(* IEC 61131-3 sources: JingjiangMoonbox/Application/Application/数据类型/系统参数/保持参数, 3 files *)

(* ---- StGrpParam_Save.st ---- *)
(*@CES
Name=StGrpParam_Save
Type=Gvl
TypeGuid=2db5746d-d284-4425-9f7f-2663a34b0ebc
Guid=f58940ec-a17f-4bea-a7e2-f076956df0df
HasDeclaration=True
HasImplementation=False
*)
{DECLARATION}
{attribute 'pack_mode' := '1'}
TYPE StGrpParam_Save :
STRUCT
	rGirth_BottomRoller							: REAL;(* 底辊周长/整机设置状态 *)
	uiNum_BottomRoller							: UINT;(* 底辊减速比分子/整机设置状态 *)
	uiDen_BottomRoller							: UINT;(* 底辊减速比分母/整机设置状态 *)

	rGirth_PrnRoller							: REAL;(* 印版周长/整机设置状态 *)
	uiNum_PrnRoller								: UINT;(* 版辊减速比分子/整机设置状态 *)
	uiDen_PrnRoller								: UINT;(* 版辊减速比分母/整机设置状态 *)

	rGirth_NetRoller							: REAL;(* 网辊周长/整机设置状态 *)
	uiNum_NetRoller								: UINT;(* 网辊减速比分子/整机设置状态 *)
	uiDen_NetRoller								: UINT;(* 网辊减速比分母/整机设置状态 *)

	rGirth_StrRoller							: REAL;(* 张带辊周长 *)
	uiNum_StrRoller								: UINT;(* 张带辊减速比分子/整机设置状态 *)
	uiDen_StrRoller								: UINT;(* 张带辊减速比分母/整机设置状态 *)

	rScrewPitch_PrnRoller_Pressure				: REAL;(* 版辊压力架丝杆节距/整机设置状态/单位mm *)
	uiNum_PrnRoller_Pressure					: UINT;(* 版辊压力电机减速比分子/整机设置状态 *)
	uiDen_PrnRoller_Pressure					: UINT;(* 版辊压力电机减速比分母/整机设置状态 *)

	rScrewPitch_NetRoller_Pressure				: REAL;(* 网辊压力架丝杆节距/整机设置状态/单位mm *)
	uiNum_NetRoller_Pressure					: UINT;(* 网辊压力电机减速比分子/整机设置状态 *)
	uiDen_NetRoller_Pressure					: UINT;(* 网辊压力电机减速比分母/整机设置状态 *)

	rScrewPitch_StrRoller_Pressure				: REAL;(* 张带辊压力架丝杆节距/整机设置状态/单位mm *)
	uiNum_StrRoller_Pressure					: UINT;(* 张带辊压力电机减速比分子/整机设置状态 *)
	uiDen_StrRoller_Pressure					: UINT;(* 张带辊压力电机减速比分母/整机设置状态 *)

	rGirth_CenterRoller							: REAL;(* 中心辊周长/整机设置状态 *)
	uiNum_CenterRoller							: UINT;(* 中心辊减速比分子/整机设置状态 *)
	uiDen_CenterRoller							: UINT;(* 中心辊减速比分母/整机设置状态 *)

	rScrewPitch_Horz							: REAL;(* 横向架丝杆节距/整机设置状态/单位mm *)
	uiNum_Horz									: UINT;(* 横向电机减速比分子/整机设置状态 *)
	uiDen_Horz									: UINT;(* 横向电机减速比分母/整机设置状态 *)

	rScrewPitch_PhotoCell						: REAL;(* 光电眼架丝杆节距/整机设置状态/单位mm *)
	uiNum_PhotoCell								: UINT;(* 光电眼电机减速比分子/整机设置状态 *)
	uiDen_PhotoCell								: UINT;(* 光电眼电机减速比分母/整机设置状态 *)

	wAI_polarity								: WORD;(* 模拟量输入极性配置 *)
		(*
		/bit0=1放料模拟量输入反向
		/bit1=1收料模拟量输入反向
		/bit2=1放牵模拟量输入反向
		/bit3=1收牵模拟量输入反向
		/bit4~bit15(保留)
		/ *)
	lrPrnLen_AmountTo							: LREAL;(* 总计印刷长度/单位:m *)
	rPrintLengthCoef							: REAL;(*印刷计长系数|*)
	alrPrnLen									: ARRAY [1..3] OF LREAL;(* A轴印长/B轴印长/总印长 *)
	alrPrnLen_Alr								: ARRAY [1..3] OF LREAL;(* 印长报警值/相对应于alrPrnLen *)
	iDelayMsec_RollerPress						: INT;(* 压辊延时/单位:ms *)

	wUwRwAxisProf								: WORD;
(*												/放料&收料轴描述 *)
(*												/bit0=TRUE,放料当前轴A轴 *)
(*												/bit1=TRUE,收料当前轴A轴 *)

	iMarkTypeId									: INT;(* 色标形式 *)
	iMarkArrangeMode							: INT;(* 标记排列形式 *)
	byTriMark_SideC								: BYTE;(* 梯形色标直边(c边) *)
	byTriMark_SideB								: BYTE;(* 梯形色标底边(b边) *)
	bySysSamplePrecision						: BYTE;(*系统采样精度			*)
	byArcFineSampleType							: BYTE;(*系统采样方式*)

	(* 时间设定 *)
	iTime_Stop									: INT;(* 停机时间/单位:s *)
	iTime_Estop									: INT;(* 急停时间/单位:s *)
	iTime_AutoAcc							: INT;(* 自动加减速时间/单位:s *)
	iTime_ManuAcc							: INT;(* 手动加减速时间/单位:s *)
	iTime_S										: INT;(* S加减速时间/单位:s *)
	iTime_PreDrvAcc_Uw								: INT;(* 预驱加速时间/10s *)
	iTime_PreDrvDec_Uw							: INT;(* 预驱减速时间/2s *)
	iTime_PreDrvAcc_Rw								: INT;(* 预驱加速时间/10s *)
	iTime_PreDrvDec_Rw							: INT;(* 预驱减速时间/2s *)
	iTime_FilmAcc								: INT;(* 料膜加速时间/8S *)
	iTime_FilmDec								: INT;(* 料膜减速时间/2S *)
	iTime_AutoDec							: INT;(*自动加减速时间|单位:s|*)
	iTime_ManuDec							: INT;(*手动加减速时间|单位:s|*)
	iTime_FastStop							: INT;(*快停时间*)
	iTime_S_End								: INT;(*S减加速时间*)
	byAutoAccDecCurve					: BYTE;(*自动加减速曲线选择|默认 按照最大直线加速度进行s处理-
																		 1：按照直线加速时间进行s处理
																		 2：按照直线加速时间全程s处理-*)

	rVel_Max									: REAL;(* 设备最大速度/单位:m/min *)
	rVel_Tar									: REAL;(* 目标速度/单位:m/min *)
	arVel_Usr									: ARRAY [1..3] OF REAL;(* 用户速度1,2,3/单位:m/min *)
	rVel_Ink									: REAL;(* 匀墨速度/单位:m/min *)
	rVel_Inch									: REAL;(* 单运行速度/单位:m/min *)
	rVel_AutoAdj								: REAL;(* 自动修正速度/单位:m/min *)
	rVel_ManuAdj_Corse							: REAL;(* 手动粗调速度/单位:m/min *)
	rVel_ManuAdj_Fine							: REAL;(* 手动细调速度/单位:m/min *)
	rVel_RapidAdj								: REAL;(* 快速调版速度/单位:m/min *)
	rVel_HorzdAdj								: REAL;(* 横向调版速度/单位:mm/s *)

	rDiamAlarm_Uw								: REAL;(* 放料报警卷径 *)
	rGirth_AxiaA_Uw								: REAL;(* 放料A轴周长 *)
	rGirth_AxiaB_Uw								: REAL;(* 放料B轴周长 *)
	arKpid_Uw									: ARRAY [1..3] OF REAL;(* 放料pid比例 *)
	rGirth_Uw									: REAL;(* 放料周长 *)
	uiNum_Uw									: UINT;(* 放料减速比-电机转数 *)
	uiDen_Uw									: UINT;(* 放料减速比-负载转数 *)
	rTaper_Uw									: REAL;(* 放料锥度 *)
	rAI_med_Uw									: REAL;(* 放料摆臂模拟量中位 *)
	byDiamMeasureTypeId_Uw						: BYTE;(* 放料卷径测量类型 *)
	byAIType_Uw									: BYTE;(* 放料摆臂类型/初始值0 *)
	byCoef_stiffen_Uw							: BYTE;(* 放料拉料系数|10 *)

	adwEnc_AxisALocation_Uw						: ARRAY [0..1] OF DWORD;(* 放料A轴定位位置/索引通过BOOL_TO_INT(xCutterOnTop_#w)来访问 *)
	adwEnc_AxisALocation_MinDiam_Uw				: ARRAY [0..1] OF DWORD;(* 放料A轴最小径位置/索引通过BOOL_TO_INT(xCutterOnTop_#w)来访问 *)
	adwEnc_AxisBLocation_Uw						: ARRAY [0..1] OF DWORD;(* 放料B轴定位位置/索引通过BOOL_TO_INT(xCutterOnTop_#w)来访问 *)
	adwEnc_AxisBLocation_MinDiam_Uw				: ARRAY [0..1] OF DWORD;(* 放料B轴最小径位置/索引通过BOOL_TO_INT(xCutterOnTop_#w)来访问 *)
	iRatedRpm_Uw								: INT;(* 放料电机额定转速/1500r/min *)
	iRatedFreq_Uw								: INT;(* 放料电机额定频率/50HZ *)
	iUpperFreq_Uw								: INT;(* 放料电机上限频率/100HZ *)
	xDiamMeasureAutomatic_Uw					: BOOL;(* 放料卷径自动测量标志/FALSE *)
	xCutUseReflectionSensor_Uw					: BOOL;(* 放料采用弧面检测方式标志,TRUE标识有效/FALSE *)
	xMultAxisParaEn_Uw							: BOOL;(* 放料AB轴单独参数-卷径测量/FALSE *)
	xFlag_CCW_AfterCutted_Uw					: BOOL;(* 裁切后放料轴反转/TRUE *)
	iPreRevLenth_MM_Cutted_Uw					: INT;(* 放料轴裁切反转距离/初始值1000 *)
	iPreRevVel_RPM_Cutted_Uw					: INT;(* 放料轴裁切反转转速/初始值80 *)
	xPreCutOneBtn_Uw							: BOOL;(* 放料接料准备使用单输入标志/FALSE *)
	rCoefCut_FilmVolPerimeter_Uw				: REAL;(* 放料裁切系数/1.5 *)
	xDiaEstEn_Uw								: BOOL;(* 放料卷径估计使能/FALSE *)
	rEstiDia_Uw									: REAL;(* 预估卷径值/300mm *)
	rEstiThickness_Uw							: REAL;(* 预估料膜厚度值/0.02mm *)
	byDelayTime_DiaCompensateWhenCutDne_Uw		: BYTE;(* 裁切后卷径补偿介入时间/10s *)
	uiPiDelay_Uw								: UINT;(* 裁切后放料PI延迟时间/1000ms *)

	xUseRadCompensate_Uw						: BOOL;(* 放料翻转架补偿使能标志/FALSE *)
	xConfirmRad0_Uw								: BOOL;(* 放料确认弧度0标志/FALSE *)
	dwAxisAabsPos_0Rad_Uw						: DWORD;(* 放料A轴翻转架0度的绝对位置/翻转架中心作为坐标系0点/0 *)
	dwAxisBabsPos_0Rad_Uw						: DWORD;(* 放料B轴翻转架0度的绝对位置/翻转架中心作为坐标系0点/0 *)
	(*											/ALTMA的放料架结构 *)
	rDiam_Tower_Uw								: REAL;(* 放料翻转架的直径/1000mm *)
	rDiam_NextRoller_Uw							: REAL;(* 放料翻转架下个辊的直径/100mm *)
	rXPos_NextRoller_Uw							: REAL;(* 放料翻转架下个辊的X位置/232.5mm/翻转架中心作为坐标系0点 *)
	rYPos_NextRoller_Uw							: REAL;(* 放料翻转架下个辊的Y位置/1052mm/翻转架中心作为坐标系0点 *)
	xTowerDir_Uw								: BOOL;(* 翻转架和绝对位置方向控制/FALSE *)
	(*2022.5.17.121911 放料翻转架补偿算法优化后增加的变量|13bytes|2023.8.17.161013*)
	rDiam_DeflectorRollPos_Uw				: REAL;(*翻料架的导向辊圆心运动直径|距离翻转架圆心=该值/2|mm*)
	rDiam_DeflectorRoller_Uw				: REAL;(*翻料架上导向辊的直径|mm*)
	xMultAxisPosEn_Uw							: BOOL;(* 放料定位位置单独参数-绝对值编码器/FALSE *)
	byInitialSpd_Stiffen_Uw						: BYTE;(* 放料拉料初始速度/10r/min *)
	(*											/ 2021.11.5.174244 *)
	rFilmLen_UnwindToPU1						: REAL;(*放料裁切点到1U的料膜距离|单位:mm|*)
	rFilmLen_NotAdjFront						: REAL;(*裁切点前不调整的料长|单位:mm|*)
	rFilmLen_NotAdjBack							: REAL;(*裁切点后不调整的料长|单位:mm|*)
	rFilmLen_BetweenImpressPoints				: REAL;(*两个压印点之间的料长|单位:mm|*)

	rDiamAlarm_Rw								: REAL;(* 收料报警卷径 *)
	rGirth_AxiaA_Rw								: REAL;(* 收料A轴周长 *)
	rGirth_AxiaB_Rw								: REAL;(* 收料B轴周长 *)
	arKpid_Rw									: ARRAY [1..3] OF REAL;(* 放料pid比例 *)
	rGirth_Rw									: REAL;(* 收料周长 *)
	uiNum_Rw									: UINT;(* 收料减速比-电机转数 *)
	uiDen_Rw									: UINT;(* 收料减速比-负载转数 *)
	rAI_med_Rw									: REAL;(* 收料摆臂模拟量中位 *)
	byAIType_Rw									: BYTE;(* 收料摆臂类型/初始值0 *)
	byCoef_stiffen_Rw							: BYTE;(* 收料拉料系数|10 *)
	xRsv										: BOOL;
	adwEnc_AxisALocation_Rw						: ARRAY [0..1,0..1] OF DWORD;(* 收料A轴定位位置/一维索引通过BOOL_TO_INT(xCutterOnTop_Rw)/二维索引[0]表示3吋纸芯,[1]表示6吋纸芯 *)
	adwEnc_AxisBLocation_Rw						: ARRAY [0..1,0..1] OF DWORD;(* 收料B轴定位位置/一维索引通过BOOL_TO_INT(xCutterOnTop_Rw)/二维索引[0]表示3吋纸芯,[1]表示6吋纸芯 *)
	rTaper_begin_Rw								: REAL;(* 锥度起始值-收料 *)
	rTaper_end_Rw								: REAL;(* 锥度结束值-收料 *)
	rDiam_taper_begin_Rw						: REAL;(* 锥度起始直径-收料 *)
	rDiam_taper_end_Rw							: REAL;(* 锥度结束直径-收料 *)
	iRatedRpm_Rw								: INT;(* 收料电机额定转速/默认1500 *)
	iRatedFreq_Rw								: INT;(* 收料电机额定频率/默认50 *)
	iUpperFreq_Rw								: INT;(* 收料电机上限频率/默认100 *)
	rGirth_3inch_Rw								: REAL;(* 收料3寸周长/默认300 *)
	rGirth_6inch_Rw								: REAL;(* 收料6寸周长/默认600 *)
	xPreCutOneBtn_Rw							: BOOL;(* 收料接料准备使用单输入标志/默认FALSE *)
	rCoefCut_FilmVolPerimeter_Rw				: REAL;(* 收料裁切系数/0.5 *)
	xDiaEstEn_Rw								: BOOL;(* 收料卷径估计使能/默认FALSE *)
	rEstiDia_Rw									: REAL;(* 预估卷径值/默认300mm *)
	rEstiThickness_Rw							: REAL;(* 预估料膜厚度值/默认0.02mm *)
	byDelayTime_DiaCompensateWhenCutDne_Rw		: BYTE;(* 裁切后卷径补偿介入时间/默认10s *)
	xUseAbsEncEn_Rw								: BOOL;(* 收料使用绝对值编码器标志/默认FALSE *)
	xMultAxisPosEn_Rw							: BOOL;(* 收料定位位置单独参数-绝对值编码器/默认FALSE *)
	byInitialSpd_Stiffen_Rw						: BYTE;(* 收料拉料初始速度/10r/min *)

	rDiamCurAxis_Uw								: REAL;(* 放料当前卷径 *)
	rDiamCurAxis_Rw								: REAL;(* 收料当前卷径 *)

	rGirth_If									: REAL;(* 放牵周长 *)
	uiNum_If									: UINT;(* 放牵减速比-电机转数 *)
	uiDen_If									: UINT;(* 放牵减速比-负载转数 *)
	rTaper_If									: REAL;(* 放牵锥度 *)
	byAIType_If									: BYTE;(* 放牵摆臂类型/初始值0 *)
	rAI_med_If									: REAL;(* 放牵摆臂模拟量中位 *)
	arKpid_If									: ARRAY [1..3] OF REAL;(* 放牵pid/2021.11.18.201839 *)
	iRatedRpm_If								: INT;(* 放牵电机额定转速/1500rpm *)
	iRatedFreq_If								: INT;(* 放牵电机额定频率/50HZ *)
	iUpperFreq_If								: INT;(* 放牵电机上限频率/100HZ *)
	xInchNegative_If							: BOOL;(* 放牵单运行反向/FALSE *)
	iInchVel_If									: INT;(* 放牵单运行速度/10m/min *)

	rGirth_Of									: REAL;(* 收牵周长 *)
	uiNum_Of									: UINT;(* 收牵减速比-电机转数 *)
	uiDen_Of									: UINT;(* 收牵减速比-负载转数 *)
	rTaper_Of									: REAL;(* 收牵锥度 *)
	byAIType_Of									: BYTE;(* 收牵摆臂类型/初始值0 *)
	rAI_med_Of									: REAL;(* 收牵摆臂模拟量中位 *)
	arKpid_Of									: ARRAY [1..3] OF REAL;(* 收牵pid/2021.11.18.202112 *)
	iRatedRpm_Of								: INT;(* 收牵电机额定转速/1500rpm *)
	iRatedFreq_Of								: INT;(* 收牵电机额定频率/50HZ *)
	iUpperFreq_Of								: INT;(* 收牵电机上限频率/100HZ *)
	xInchNegative_Of							: BOOL;(* 收牵单运行反向/FALSE *)
	iInchVel_Of									: INT;(* 收牵单运行速度/10m/min *)

(*2025.8.4.144213|原dwExtBitCtlFlag变量-改为BIT型--*)
	xSwitch_Change_CutterOnTop_HMI_Uw			: BIT;(*放料上下裁切换-界面按钮bit2*)
	xSwitch_Change_CutterOnTop_HMI_Rw			: BIT;(*收料上下裁切换-界面按钮bit3*)
	xCancelTenEn								: BIT;(*取消张力规划使能开bit10*)
	xEn_DualParam_AbsEncLocation_Uw				: BIT;(*bit11: 放料编码器方式下定位使用多轴使能|2021.5.7.111434|Liu.yt*)
	xEn_DualParam_AbsEncLocation_Rw				: BIT;(*bit12: 收料编码器方式下定位使用多轴使能|2021.5.7.111434|Liu.yt*)
	xFlag_AxisABParaFroDiaMea_Uw				: BIT;(*放料自动卷径分轴标志*)
	xSwitchTension_If							: BIT;(*bit6 放牵张力算法切换/FALSE *)
	xSwitchTension_Of							: BIT;(*bit7 收牵张力算法切换/FALSE *)
	xEnFeedLimitWarnFlag						: BIT;(*bit5 牵引速度限制提示使能位*)
	xSwitch_AxisLocaltion_DualParam_Uw			: BIT;(*放料绝对值编码器定位双轴参数开关|原bit11*)
	xSwitch_AxisLocaltion_DualParam_Rw			: BIT;(*收料绝对值编码器定位双轴参数开关|原bit12*)
	dwExtBitCtlFlag								: DWORD;(*扩展位控制标志|2019.1.25.143212|
													*.bit0: 放料自动卷径是否分轴来作?|FALSE默认一起|TRUE表示ab轴分开||
													*.bit1: 一键开机使能标志||
													*.bit2: 放料上下裁控制开关(区分于xCutterOnTop_Uw|)|2019.3.28.092931|补充遗漏||
													*.bit3: 收料上下裁控制开关(区分于xCutterOnTop_Rw|)|2019.3.28.092931|补充遗漏||
													Deprecated@2019.8.13.115259|*.bit4: 超声波检测使能|2019.3.23.154021||2019.3.28.092949|纠正错误||
													*.bit5: 牵引速度限制提示使能位|2019.4.18.135612|xie.gc||
													*.bit6: 放牵算法切换开关|@2019.8.1.091703|
													*.bit7: 收牵算法切换开关|@2019.8.1.091703|
													*.bit8: 放料前馈使能位|@2019.8.8.162527|xie.gc|
													*.bit9: 收料前馈使能位|@2019.8.8.162527|xie.gc|
													*.bit10: 取消张力规划使能开|2019.10.14.152513|niu.j|
													*.bit11: 放料编码器方式下定位使用多轴使能|2021.5.7.111434|Liu.yt|
													*.bit12: 收料编码器方式下定位使用多轴使能|2021.6.1.093832|Liu.yt|
													ALTMA增加了上下裁刀是否配置标志
													*.bit13: |2021.7.17.142536 放料上裁刀开启|Liu.yt|
													*.bit14: |2021.7.17.142536 放料下裁刀开启|Liu.yt|
													*.bit15: |2021.7.17.142536 收料上裁刀开启|Liu.yt|
													*.bit16: |2021.7.17.142536 收料下裁刀开启|Liu.yt|
													*.bit17: 2022.4.6.130956\翻料架打开控制位|
													|*)

	byTaperCtlMode_Uw							: BYTE;(*锥度调整方式*)
	byTaperCtlMode_Rw							: BYTE;(*锥度调整方式*)
	(*2022.4.14.094534 收放料自动接料|21BYTES*)
	xAutomaticCutEn_Uw							: BOOL;(*放料自动裁切使能|*)
	byAutoMaticCutMode_Uw						: BYTE;(*放料自动裁切模式|0 按照剩余米数
																	 |1 按照剩余卷径*)
	uiAutoMaticCutMeters_Uw						: UINT;(*自动裁切米数|m*)
	uiAutoMaticCutDia_Uw						: UINT;(*自动裁切卷径|*)

	xAutomaticCutEn_Rw							: BOOL;(*收料自动裁切使能|*)
	byAutoMaticCutMode_Rw						: BYTE;(*收料自动裁切模式|0 按照计米长度-在上次接料完成后启动
															         |1 按照放料裁切后整机长度-在放料接料完成后启动
																     |2 按照当前卷径-在上次接料完成后启动*)
	uiAutoMaticCutMeters_Rw						: UINT;(*自动裁切米数|m*)
	uiAutoMaticCutDia_Rw						: UINT;(*自动裁切卷径|*)
	byLenth_Machine								: BYTE;(*整机长度|m*)
	rDia_PaperRoller_Uw							: REAL;(*纸筒直径|mm*)
	rFilmThickNess								: REAL;(*料膜厚度|mm*)
	(*放料|*)
	rDiamTaper_Begin_Uw							: REAL;(*放料起始锥度对应卷径|*)
	rDiamTaper_End_Uw							: REAL;(*放料结束锥度对应卷径|*)
	rTaper_Begin_Uw								: REAL;(*锥度起始|放料|*)
	rTaper_End_Uw								: REAL;(*锥度结束|放料|*)

	(*放牵|*)
	rTaper_Begin_If								: REAL;(*锥度起始|放牵|*)
	rTaper_End_If								: REAL;(*锥度结束|放牵|*)
	(*收牵|*)
	rTaper_Begin_Of								: REAL;(*锥度起始|收牵|*)
	rTaper_End_Of								: REAL;(*锥度结束|收牵|*)

	xStep_Fast:BOOL;
	rStep_Fast:REAL;
	rStep_Little:REAL;
(*增加收放料收放牵锥度单位切换|支持%、N、mpa|104bytes*)
	byTaperUnit_Uw								: BYTE;(*放料锥度单位|默认%*)
	rPercentMatchN_Uw							: REAL;(*放料百分比-单位是N的对应|确认的值*)
	rN_Uw										: REAL;(*放料牛顿值|确认的值*)
	rPercentMatchMpa_Uw							: REAL;(*放料百分比-单位是Mpa的对应|确认的值*)
	rMpa_Uw										: REAL;(*放料兆帕值|确认的值*)

	byTaperUnit_Rw								: BYTE;(*收料锥度单位|默认%*)
	rPercentMatchN_Rw							: REAL;(*收料百分比-单位是N的对应|确认的值*)
	rN_Rw										: REAL;(*收料牛顿值|确认的值*)
	rPercentMatchMpa_Rw							: REAL;(*收料百分比-单位是Mpa的对应|确认的值*)
	rMpa_Rw										: REAL;(*收料兆帕值|确认的值*)

	byTaperUnit_If								: BYTE;(*放牵锥度单位|默认%*)
	rPercentMatchN_If							: REAL;(*放牵百分比-单位是N的对应|确认的值*)
	rN_If										: REAL;(*放牵牛顿值|确认的值*)
	rPercentMatchMpa_If							: REAL;(*放牵百分比-单位是Mpa的对应|确认的值*)
	rMpa_If										: REAL;(*放牵兆帕值|确认的值*)

	byTaperUnit_Of								: BYTE;(*收牵锥度单位|默认%*)
	rPercentMatchN_Of							: REAL;(*收牵百分比-单位是N的对应|确认的值*)
	rN_Of										: REAL;(*收牵牛顿值|确认的值*)
	rPercentMatchMpa_Of							: REAL;(*收牵百分比-单位是Mpa的对应|确认的值*)
	rMpa_Of										: REAL;(*收牵兆帕值|确认的值*)
	rDiamCurAxis_Uw2							: REAL;

	(*2025.8.9.142811增加*)
	xUseBtn_Linkage							: BIT;(*联动使用按钮/FALSE:开关|原wCtlSwitchRef.5*)
	xSwitch_WaitFilmLengthEn				: BIT;(*开机等料长|原原wCtlSwitchRef.4*)
	xSwitch_WaitFilmLengthEn_From1st		: BIT;(*开机等首色料长|原原wCtlSwitchRef.13*)
	xSwitch_GiveupHeaderEn					: BIT;(*让料头|原wCtlSwitchRef.15*)
	xSwitch_Alarm_Arc						: BIT;(*套色报警开关|wCtlSwitchRef.0*)
	xSwitch_InkRollerSolenoid_Use3			: BIT;(*递墨辊三档有效标志|原wCtlSwitchRef.9*)
	xBitRsv6: BIT;
	xBitRsv7: BIT;
//2025.12.30.215929注意新增变量了，参数不统一了
	byIn_outFeed_ThresCoff							: BYTE;(*断料保护牵引判断阀值|原LREAL型，改为BYTE吧*)
//2026.1.9.160446这里替代一下先防止数据大小变化
//	byBitRsv: BYTE;
	byBitRsv1: BYTE;
	(*2025.10.14.134703先把这个屏蔽了，直接用bit类型吧|NIU.J
	wCtlSwitchRef							: WORD;(*整机控制开关描述|
													*.bit0: 套色报警开关
													*.bit1: 波门锁|根据色组来更新
													*.bit2: 整机纵向自动| 2018.3.23.145133| han.dp|
													*.bit3: 整机横向自动| 2018.3.23.145153| han.dp|
													*.bit4: 开机等料长\2018.5.27.153018|
													*.bit5: han.dp\2018.6.19.172042\联动采用非两档开关|
													*.bit6: 2018.7.13.081355\使能标准3''6''纸管选择|TRUE按标准纸管走 FALSE按屏幕输入走|
													*.bit7: 2018.7.3.194246\色组单独减速比设置|
													*.bit8: 2018.7.23.143553\刮刀使能开关|
													*.bit9: 2018.7.28.102401\递墨辊三档有效标志|(TRUE有效)|
													*.bit10: 2018.8.13.101345\预加热印刷使能|
													*.bit11: 排风限制热风使能|
													*.bit12: 2018.8.15.082652\放料表印选择\默认FALSE=里印|
													*.bit13: 2018.8.15.082652\收料表印选择\默认FALSE=里印|
													*.bit14: 2022.4.6.140140排风限制开机使能
													|*)
													*)

	wCtl_Pressure_Up_Dn							: WORD;
												(*
												bit0：自动合压-进入印刷状态后自动合压
												bit1：急停直接离压/FALSE急停不动作，复位离压
												bit2：裁切避让胶带使能
												bit3：裁切避让胶带外触发标志/内触发需要计算裁切切点到1色料长
												bit4：停机自动匀墨
												bit5：压力电机维持使能
												bit6：点位运动电机维持使能
												*)
	rLength_AvoidancePoint_To_1u_mm				: REAL;//避让胶带检测点到1色的距离

	rFilmThick_Confirm							: REAL;
	rFilmThick_Manu								: REAL;

	lrDistanceOfLimitTo_MEdge_MM				: LREAL;//限位距离边缘的距离,单位 ： mm
//秦华带长相关功能标志
	xLength_BandLen_Check						: BOOL;(*手动检测带长*)
	rLength_Band_Confirm						: REAL;(* 带长/整机设置状态,需要同步到每个色组的检测带长 *)
	xLength_BandLen_Sync						: BOOL;(*自动同步带长*)
	rLength_HeightStandard						: REAL;(*整机同步带长的标准纵向高度值*)
	rLength_Width								: REAL;(*版辊张带辊横向差值*)
	rLength_Printing : REAL;		//系统印长
//2024.12.11.135813 | 增加印版辊速度、网辊速度、张带速度		12字节
	rVel_Press_Prn:REAL;
	rVel_Press_Net:REAL;
	rVel_Press_Str:REAL;
	rPressure_Tar : REAL;
//2025.02.27.200725 | 增加收放料小卷径补偿		18字节
	xSmallDiaMulEn_UW						: BOOL;//:= FALSE;
	iSmallDiaMulSa_UW						: INT;//:=200;(*进入该方式的启动卷径|大卷径*)
	iSmallDiaMulEd_UW						: INT;//:=100;(*结束的卷径|写死为最小卷径*)
	iSmallDiaMulSa_Coeff_UW					: INT;//:=100;(*系数|单位%*)
	iSmallDiaMulEd_Coeff_UW					: INT;//:=300;(*系数|单位%*)

	xSmallDiaMulEn_RW						: BOOL;//:= FALSE;
	iSmallDiaMulSa_RW						: INT;//:=200;(*进入该方式的启动卷径|大卷径*)
	iSmallDiaMulEd_RW						: INT;//:=100;(*结束的卷径|写死为最小卷径*)
	iSmallDiaMulSa_Coeff_RW					: INT;//:=100;(*系数|单位%*)
	iSmallDiaMulEd_Coeff_RW					: INT;//:=300;(*系数|单位%*)
//	2025.02.28.092405 /增加色组间加热控制的两档位 		4字节
	rVel_Temp_I								: INT;//:=30;
	rVel_Temp_II							: INT;//:=60;
	rBandLengthNotAdjArea					: REAL;
	rVel_NetReturn : REAL;

	iVelSa_ScraperRun						: INT;
	iVolt_ScraperMin						: INT;(*刮刀变频最小电压|2018.7.25.121151|*)
	iVolt_ScraperMax						: INT;(*刮刀变频最大电压|2018.7.25.121151|*)
	lrRatedRpm_Scraper						: LREAL;(*刮刀变频额定转速|*)
	lrRatedFreq_Scraper						: LREAL;(*刮刀变频额定频率|*)
	lrUpperFreq_Scraper						: LREAL;(*刮刀变频上限频率|*)
	lrLowerFreq_Scraper						: LREAL;(*刮刀变频下限频率|*)
	rMaxFreq_Scraper						: REAL;(*刮刀变频最大频率|*)
	rMinFreq_Scraper						: REAL;(*刮刀变频最小频率|*)

	lrCoeff_Scraper							: LREAL;(*刮刀变频速度系数|*)
	iNum_ScraperMotor						: INT;(*刮刀电机减速比分子numerator*)
	iDen_ScraperMotor						: INT;(*刮刀频率分母denominator*)
	iRatio_ScraperContrastToPrintRoller		: INT;(*刮刀相对版转速的对应比*)
	iDelayMsec_Heat							: INT;(*加热延时时间|*)
	iDelayMsec_HeatBlower					: INT;(*热风延时时间|*)
	iDelayMsec_ExhPowerMode					: INT;(*排风模式切换时间|*)

	(*张力优化算法2025.7.3.175755*)
	rR_K_LQR_Uw												: REAL;
	rN_LQR_Uw												: REAL;
	rR_K_MinBeat_Uw											: REAL;
	iN_MinBeat_Uw											: INT;
	xUseAntiNotch_Uw										: BOOL;(*套色使用陷波器@*)
	rWn_Uw													: REAL;(*陷波中心频率 rad/s*)
	rBw_Uw													: REAL;(*陷波宽度 rad/s*)
	rDp_Uw													: REAL;(*陷波深度 dB*)
	xUseIMatrix_rX_DARE_Uw									: BOOL;(*使用单位矩阵否则使用的是特定卷径的收敛值*)
	rKc_Uw													: REAL;(*补偿系数*)
	rKc_Uw_AccDec											: REAL:=0.08;(*加减速时候输出系数@必须为负值*)
	uiUseTime_Diam_Min_Uw									: UINT;(*使用时变的最小卷径|mm@2024.05.14.080937*)
	xUseTime_b1_Uw											: BOOL;(*有效则b1随卷径实时变化-不实时变化则使用b1_0@2024.05.14.080937*)
	xUseDiam_LowPass_Uw										: BOOL;(*使用低通滤波后的卷径*)
	rWc_LowPass_Diam_Uw										: REAL;(*放料卷径低通截止频率@2024.7.11.152456*)
	xUseIfVel_Uw											: BOOL;(*使用放牵速度|放料张力算法以及原来的前馈@2024.8.21.165317*)

	rR_K_LQR_Rw												: REAL;
	rN_LQR_Rw												: REAL;

	rR_K_MinBeat_Rw											: REAL;
	iN_MinBeat_Rw											: INT;

	xUseIMatrix_rX_DARE_Rw									: BOOL;(*使用单位矩阵否则使用的是特定卷径的收敛值*)
	rKc_Rw_AccDec											: REAL:=0.08;(*加减速时候输出系数@必须为负值*)
	uiUseTime_Diam_Min_Rw									: UINT;(*使用时变的最小卷径|mm@2024.05.14.080937*)
	xUseTime_b1_Rw											: BOOL;(*有效则b1随卷径实时变化-不实时变化则使用b1_0@2024.05.14.080937*)
	rKc_Rw													: REAL;(*补偿系数*)
	byKalmanFilterType_Rw									: BYTE;(*收料张力估计时卡尔曼滤波类型选择*)

	(*收料张力算法使能标志@2024.7.15|11bytes*)
	xTensionCompensateEn_Rw									: BOOL;(*张力补偿算法使能*)
	xTensionCompensateEn_RwCut								: BOOL;(*收料裁切使用张力补偿使能*)
	xUseDiam_LowPass_Rw										: BOOL;(*使用低通滤波后的卷径*)
	rWc_LowPass_Diam_Rw										: REAL;(*收料卷径低通截止频率*)
	rWuCompensate_Rw										: REAL;(*补偿的转速(R/MIN)|计算的*)
	rWuCompensate_Act_Rw									: REAL;(*补偿的转速(R/MIN)|实际使用的*)

	xUseOfVel_Rw											: BOOL;(*使用收牵速度|收料张力算法以及原来的前馈@2024.8.21.165317*)
(*	abyReserved_TensionCtl_Rw								: ARRAY [1..1] OF BYTE;*)
											(*xUseOfVel_Rw|0*)
											(*xTensionCompensateEn_Rw-->xTensionCompensateEn_RwCut|16->1*)
	(*收放料新的pid算法标志*)
	xPidType_If_New							: BOOL;
	xPidType_Of_New							: BOOL;
(*2025.7.3.175755开始增加内容*)
	byKalmanFilterType_Uw:BYTE;(*放料张力估计时卡尔曼滤波类型选择@=0 Kalman_CycDis_BeiRen/Kalman_CycDis_test
																 @=1 Youla_Kalman
																 @=2 ExtendKalman
																 @=3 UnExtendKalman*)
	byStructParanInitEn_Uw									: BYTE;(*初始化使能标志@按照定义顺序/.0 初始化第一个结构体。以此类推！@顺序按照KS_InitTensionCtl_StructParam定义*)
	byStructParanInitEn_Rw									: BYTE;(*初始化使能标志@按照定义顺序/.0 初始化第一个结构体。以此类推！@顺序按照KS_InitTensionCtl_StructParam定义*)

	byNeedAutomaticCut_UwRw									: BYTE;	(*打开自动裁切使能提示标志@按系区分*)
	(*2025.7.3.175755增加*)
	iCutDneResetPidMultiple_Uw								: INT;(*裁切后PID放大倍数*)
	iCutDneResetPidMultiple_Rw								: INT;(*裁切后PID放大倍数*)
	iCutDneResetPidRemainTime_Uw							: INT;
	iCutDneResetPidRemainTime_Rw							: INT;
	iCutDneResetPidToDefaultTime_Uw							: INT;
	iCutDneResetPidToDefaultTime_Rw							: INT;
	xUseAbsEncoder_Uw										: BOOL;(*放料编码器方式定位*)
	xUseAbsEncoder_Rw										: BOOL;(*收料编码器方式定位*)
	uiPreStopDelayTime_ms									: UINT:=100;(*预驱停止延迟时间@100ms*)
	dwAbsEnCodeResolution_Uw					: DWORD;(* 放料绝对值编码器分辨率/8388608 *)
	dwAbsEnCodeResolution_Rw					: DWORD;(* 收料绝对值编码器分辨率/8388608 *)
	xUseFollow_1U_V_UwCut					: BOOL;(*使用放料裁切跟踪第一色方法*)
	uiMaxDia								: UINT;(*最大的卷径@mm*)
	uiInitDiam_Uw							: UINT;(*初始的卷径@mm|=0 按照200---uiMaxDia取中间值*)
	uiInitDiam_Rw							: UINT;(*初始的卷径@mm|=0 按照200---uiMaxDia取中间值*)
	xGetFilmThickNessAuto					: BOOL;(*料膜厚度获取方式*)
	rFilmThickNess_Using					: REAL;(*最终应用的料膜厚度*)
	byAlarmType_NoMaterial_Uw				: BYTE:=0;(*没料报警方式@=0 放料没料3S响铃报警
													  @=1 放料没料时候一直报警-直到按下正转\反转\接料准备*)
	xTensionCompensateEn_Uw					: BOOL;
	xTensionCompensateEn_UwCut				: BOOL;
	xUseTime_Variaition_Uw					: BOOL;(*使用时变参数标志*)
	xUseTime_Variaition_Rw					: BOOL;(*使用时变参数标志*)
	byAlarmHold_PreCut_Uw					: BYTE;
	byAlarmHold_PreCut_Rw					: BYTE;
	xCutDneResetPidEn_Uw					: BOOL;
	xCutDneResetPidEn_Rw					: BOOL;
	byMeters_UseFollow_1U_V_UwCut			: BYTE;(*裁切时跟一色*)
	byVelSa_DiamCompensate_Uw				: BYTE;
	byVelSa_DiamCompensate_Rw				: BYTE;
	xGetLenthMachine_Rw:BOOL;(*收料自动裁切获取料长使能*)
	xUseKnob_6Inch_Rw_Hmi: BOOL;(**)(*收料3-6寸使用界面旋钮@2024.04.18.182812*)
	byPrintLength_CalcCtl					: BYTE;(*控制印刷记长显示|niu.j|2019.1.25.135921||*)
	alrPrnLen_FilmVel						: ARRAY [1..3] OF LREAL;(*根据料膜速度计算记米|niu.j|2019.1.25.135921||*)
	alrPrnLen_PTPos							: ARRAY [1..3] OF LREAL;(*根据PT规划位置计算记米|niu.j|2019.1.25.135921||*)
	alrPrnLen_FilmCnt						: ARRAY [1..3] OF LREAL;(*根据幅数记米|niu.j|2019.1.25.135921||*)

	xCompensateWhenAccing_If			:BOOL:=FALSE;
	rCompensateGirthWhenAccing_If		:REAL:=0;(*补偿的值|mm*)
	xCompensateWhenAccing_Of			:BOOL:=FALSE;
	rCompensateGirthWhenAccing_of		:REAL:=0;(*补偿的值|mm*)
	byVelLimit_PerCent_IfOf				: BYTE;
	iFeedLimitWarnCoff					: INT;(*牵引调整fazhi*)
	xUseAntiNotch_If					: BOOL;
	xUseAntiNotch_Of					: BOOL;
	rWn_If								: REAL;
	rBw_If								: REAL;
	rDp_If								: REAL;
	rWn_Of								: REAL;
	rBw_Of								: REAL;
	rDp_Of								: REAL;

	(*2025.8.6.193451套色调整*)
	iWorkMode_Pid						: INT;(*1-传统pid; 2-目标pid|*)
	xFlag_Follow_1U_H						:BOOL;
	xFlag_Follow_1U_V						:BOOL;
	(*目前取值2--6|该值代表当前色不受前n个轴影响
	即为2时是解耦每个机组的前两组(第3组不受第2组影响；第4组不受第2、3组影响；第5组不受第3、4组影响*)
	byDeCoupleArcNum:BYTE;(*解耦的深度|默认先取3*)
	byDeCoupleDelayNum:BYTE;(*解耦时延拍数|默认先取18*)
	rFilmLenth_InUnit:REAL;(*色组间料长单位|m@测试先写成系参数*)
	byInitTaper_Rw: BYTE;
	rInitTaper_Hmi_Rw: REAL;
	rPressure_Max									:REAL		;(*涂布压力传感器最大标定值*)
	rHz_MainExhaust_ManuallySet						:REAL	;(*主排风设定频率*)
	byStationIdDst_VirEnc							:BYTE		;(*异站编码器目标站好*)
	iPreHotRoller_Velocity_PreHot 					:INT	;  (*预热辊额定转速*)
	rStandardFreq_HotRoller_PreHot 					:REAL	; (*预热辊额定频率*)
	rUpperFreq_HotRoller_PreHot 					:REAL	;    (*预热辊上限频率*)
	rCoeff_HotRoller_PreHot 						:REAL;        (*预热辊速度系数*)
	rGirth_HotRoller_PreHot 						:REAL	;        (*预热辊周长*)
	iPreAirHotRollTorque 							:INT;           (*预热辊转矩*)
	uiDen_HotRoller_PreHot 							:UINT	;         (*预热辊减速比分母*)
	uiNum_HotRoller_PreHot 							:UINT;         (*预热辊减速比分子*)
	iPreHotRoller_Velocity_Water 					:INT	;   (*水冷辊额定转速*)
	rStandardFreq_HotRoller_Water 					:REAL	;  (*水冷辊额定频率*)
	rUpperFreq_HotRoller_Water 						:REAL	;     (*水冷辊上限频率*)
	rCoeff_HotRoller_Water 							:REAL;         (*水冷辊速度系数*)
	rGirth_HotRoller_Water 							:REAL	;         (*水冷辊周长*)
	uiDen_HotRoller_Water 							:UINT	;          (*水冷辊减速比分母*)
	uiNum_HotRoller_Water 							:UINT;			(*水冷辊减速比分子*)
	byHotBlowerStopDelayTime 						:BYTE;		  (*热风停止延时*)
	byFreqMin_HotWind 								:BYTE	;				(*热风最小频率*)
	byFreqMax_HotWind 								:BYTE	;				(*热风最大频率*)
	byDelayTime_PressDneInPrint_If 					:BYTE		;		 (*放牵压辊延时*)
	byAxisInitPhaseTypeWhenPreRegister 				:BYTE;              	(*预套准初始位置*)
	rAdjVal_PerTime_Fine : REAL;(*手动细调调整量*)
	rAdjVal_PerTime_Coarse : REAL;(*手动粗调调整量*)
	rVel_HorzPreRegister : REAL;(*横向预套准速度*)

	rVel_Tar_9905			: REAL;
	iMicron_StepTest1_V		: INT;
	iMicron_StepTest2_V		: INT;
	R_0_RW				: REAL;
	a0_0_RW	        	: REAL;
	b1_0_RW	        	: REAL;
	Wn_0_RW	        	: REAL;
	Beta_0_RW	    	: REAL;
	l_0_RW	        	: REAL;
	K_PI_RW	        	: REAL;
	a_RW	            : REAL;
	b_RW	            : REAL;
	Ts_RW	            : REAL;
	Range_RW	        : REAL;
	Theta_RW	        : REAL;
	K_adj_RW	        : REAL;
	R_0_UW		: REAL	;
	a0_0_UW     : REAL 	;
	b1_0_UW     : REAL 	;
	Wn_0_UW     : REAL 	;
	Beta_0_UW   : REAL 	;
	l_0_UW      : REAL 	;
	K_PI_UW     : REAL 	;
	a_UW        : REAL 	;
	b_UW        : REAL 	;
	Ts_UW       : REAL 	;
	Range_UW    : REAL 	;
	Theta_UW    : REAL 	;
	K_adj_UW    : REAL 	;

(*部分开关变量2025.8.8.152013*)
	xSwitch_StartUp					: BIT;(*一键开机*)
	xSwitch_RollOver				: BIT;(*翻料架开关*)
	(*新增变量-开始-2025.08.11.135045*)
	xHor_Goal_Flag : BOOL;(*横向目标值标志*)
	xHor_PreRegist_Flag : BOOL;(*横向重复值标志*)
	xEnaTestARC_Ink : BOOL;(*空转测试使能*)
	xHorLimit : BOOL; (*限位定义修改为左右|默认是正反转*)
	xHorManuCtrl:BOOL; (*界面横向手动修正功能*)
	(*新增变量-结束-2025.08.11.135057*)

(*原用户基础工艺开关控制位直接用BIT吧，不用dwCtlBits_UnitBaseCraft了--
通讯改为共用体吧*)
(*bit0-bit31--2025.8.13.100117*)
	xSwitch_ScraperAuto_If					: BIT;(*刮刀手自动-bit0*)
	xSwitch_ScraperOn_If					: BIT;(*刮刀开关bit1*)
	xInterver_ScraperRun_If					: BIT;(*刮刀开关bit2*)
	xRsv_BIT3_If							: BIT;(*BIT3预留*)
	xSwitch_InkRollerAuto_If				: BIT;(*递墨辊手自动bit4*)
	xSwitch_InkRollerCW_If					: BIT;(*递墨辊正转bit5*)
	xSwitch_InkRollerCCW_If					: BIT;(*递墨辊反转bit6*)
	xInterver_InkRollerRun_If				: BIT;(*递墨辊运行bit7*)
	xInterver_HotWindRun_If					: BIT;(*热风1运行bit9*)
	xRsv_BIT10_If							: BIT;(*BIT10预留*)
	xRsv_BIT11_If							: BIT;(*BIT11预留*)
	xSwitch_HotWindOn_II_If					: BIT;(*热风开关bit12*)
	xInterver_HotWindRun_II_If				: BIT;(*热风1运行bit13*)
	xRsv_BIT14_If							: BIT;(*BIT14预留*)
	xRsv_BIT15_If							: BIT;(*BIT15预留*)
	xSwitch_HeatingMode_Water_If			: BIT;(*水加热开关bit16*)
	xSwitch_HeatingMode_Ele_If				: BIT;(*电加热开关bit17*)
	xSwitch_Heating_II_If					: BIT;(*加热II档bit19*)
	xSwitch_Heating_III_If					: BIT;(*加热III档bit20*)
	xRsv_BIT21_If							: BIT;(*BIT21预留*)
	xRsv_BIT22_If							: BIT;(*BIT22预留*)
	xErrReset_Scraper_If					: BIT;(*刮刀故障复位bit23*)
	xErrReset_InkRoller_If					: BIT;(*递墨故障复位bit24*)
	xErrReset_Hotwind_If					: BIT;(*热风故障复位bit25*)
	xErrReset_Hotwind_II_If					: BIT;(*热风2故障复位bit26*)
	xErrReset_ExhAir_If						: BIT;(*排风故障复位bit27*)
	xSwitch_ExhAir_If						: BIT;(*排风开关bit28*)
	xInterver_ExhAir_If						: BIT;(*排风运行bit29*)
	xRsv_BIT30_If							: BIT;(*BIT30预留*)
	xSwitch_Coolwind_If						: BIT;(*冷风开关*)

	xSwitch_PreHotAirEn								: BIT;
	xSwitch_PreHeatingEn							: BIT;

(*基础工艺开关-*)
(*原用户基础工艺开关控制位直接用BIT吧，不用dwCtlBits_UnitBaseCraft了--
通讯改为共用体吧*)
(*bit0-bit31--2025.8.13.100117*)
	xSwitch_ScraperAuto_Of					: BIT;(*刮刀手自动-bit0*)
	xSwitch_ScraperOn_Of					: BIT;(*刮刀开关bit1*)
	xInterver_ScraperRun_Of					: BIT;(*刮刀开关bit2*)
	xRsv_BIT3_Of							: BIT;(*BIT3预留*)
	xSwitch_InkRollerAuto_Of				: BIT;(*递墨辊手自动bit4*)
	xSwitch_InkRollerCW_Of					: BIT;(*递墨辊正转bit5*)
	xSwitch_InkRollerCCW_Of					: BIT;(*递墨辊反转bit6*)
	xInterver_InkRollerRun_Of				: BIT;(*递墨辊运行bit7*)
	xSwitch_HotWindOn_Of					: BIT;(*热风开关bit8*)
	xInterver_HotWindRun_Of					: BIT;(*热风1运行bit9*)
	xRsv_BIT10_Of							: BIT;(*BIT10预留*)
	xRsv_BIT11_Of							: BIT;(*BIT11预留*)
	xSwitch_HotWindOn_II_Of					: BIT;(*热风开关bit12*)
	xInterver_HotWindRun_II_Of				: BIT;(*热风1运行bit13*)
	xRsv_BIT14_Of							: BIT;(*BIT14预留*)
	xRsv_BIT15_Of							: BIT;(*BIT15预留*)
	xSwitch_HeatingMode_Water_Of			: BIT;(*水加热开关bit16*)
	xSwitch_HeatingMode_Ele_Of				: BIT;(*电加热开关bit17*)
	xSwitch_Heating_I_Of					: BIT;(*加热I档bit18*)
	xSwitch_Heating_II_Of					: BIT;(*加热II档bit19*)
	xSwitch_Heating_III_Of					: BIT;(*加热III档bit20*)
	xRsv_BIT21_Of							: BIT;(*BIT21预留*)
	xRsv_BIT22_Of							: BIT;(*BIT22预留*)
	xErrReset_Scraper_Of					: BIT;(*刮刀故障复位bit23*)
	xErrReset_InkRoller_Of					: BIT;(*递墨故障复位bit24*)
	xErrReset_Hotwind_Of					: BIT;(*热风故障复位bit25*)
	xErrReset_Hotwind_II_Of					: BIT;(*热风2故障复位bit26*)
	xErrReset_ExhAir_Of						: BIT;(*排风故障复位bit27*)
	xSwitch_ExhAir_Of						: BIT;(*排风开关bit28*)
	xInterver_ExhAir_Of						: BIT;(*排风运行bit29*)
	xRsv_BIT30_Of							: BIT;(*BIT30预留*)
	xSwitch_Coolwind_Of						: BIT;(*冷风开关*)
(*基础工艺开关-*)
(*刮刀递墨一控多相关参数*)
	rHz_Scraper_ManuallySet				: REAL;(*刮刀手动频率*)
	(*新增变量-开始|wang.nt|2025.08.12.163420*)
	xLostPressure:BOOL;(*气压低报警|不允许开机*)
	xPrnRollerLoose_AtLeast1:BOOL;(*至少1色夹板报警|不允许开机*)
	xbrakeResistanceTempHigh_AtLeast1:BOOL;(*至少1色制动电阻温度过高*)
	(*新增变量-结束|wang.nt|2025.08.12.163420*)

(*2025.8.13.114803新增递墨参数*)
	iRatedRpm_InkRoller						: INT;(*递墨辊变频额定转速|*)
	iRatedFreq_InkRoller					: INT;(*递墨辊变频额定频率|*)
	iUpperFreq_InkRoller					: INT;(*递墨辊变频上限频率|*)
	iVel_InkRollerMin						: INT;(*递墨辊变频最小频率对应最小速度|*)
	iFrq_InkRollerMin						: INT;(*递墨辊变频最小频率|*)
	iVel_InkRollerMax						: INT;(*递墨辊变频最大频率对应的最大速度|*)
	iFrq_InkRollerMax						: INT;(*递墨辊变频最大频率|*)
	rCoeff_InkRoller						: REAL;(*递墨辊变频速度系数|*)
	iVelSa_InkRollerRun						: INT;(*递墨辊可以运行的起始速度|2022.5.19.130612*)

(*2025.8.13.114803新增递墨参数*)
	rHz_InkRoller_ManuallySet			: REAL;(*刮刀手动频率*)
	(*新增变量-开始|wang.nt|2025.08.12.163420*)
	xBtn_ResetAlarm:BOOL;(*按钮被按下*)
	xFlag_PhaseRead:BOOL;(*读取装版相位*)
	iOneKeySwitchOn_IdGSE: INT;(*当前系处于一键开机*)
	iMotionCtlErrCode:INT;(*错误*)
	xTips_ExhausLimitStart:BOOL;(*排风限制开机*)
	xHorzMotorAlarmAtLeastOne:bool;(*横向电机报警*)
	(*新增变量-结束|wang.nt|2025.08.12.163420*)

	xWorkMode_RollerPress					: BOOL;(*压辊顺序; TRUE从前到后; FALSE从后到前|*)
	//结构体定义
	astStTimeSet_DnCut_UpCut_Uw					: ARRAY [0..1] OF StTimeSet_DnCut_UpCut;(* 放料端的裁切时间集/BOOL_TO_INT(xCutterOnTop_Uw)做索引访问 *)
	astStTimeSet_DnCut_UpCut_Rw					: ARRAY [0..1] OF StTimeSet_DnCut_UpCut;(* 收料端的裁切时间集/BOOL_TO_INT(xCutterOnTop_Rw)做索引访问 *)
	astStStdVolParam_DnCut_UpCut				: ARRAY [0..1] OF StStdVolParam_DnCut_UpCut;(* 卷径测量参数集/BOOL_TO_INT(xCutterOnTop_Uw)做索引访问 *)
	stModelParam_Uw								: Initial_Model_Parameters;(*放料模型初始参数@50bytes*)
	stInvariant_Parameters_Uw					: Invariant_Parameters;(*放料张力算法系统参数@30bytes*)
	stPI_Parameters_Uw							: PI_Parameters;(*控制器pi参数@20bytes|用于稳速*)
	stPI_Parameters_Uw_AccDec					: PI_Parameters;(*控制器pi参数@20bytes|2024.05.13.180942 增加一组加减速的控制参数*)

	stModelParam_Rw								: Initial_Model_Parameters;(*放料模型初始参数@50bytes*)
	stInvariant_Parameters_Rw					: Invariant_Parameters;(*放料张力算法系统参数@30bytes*)
	stPI_Parameters_Rw							: PI_Parameters;(*控制器pi参数@20bytes|用于稳速*)
	stPI_Parameters_Rw_AccDec					: PI_Parameters;(*控制器pi参数@20bytes|2024.05.13.180942 增加一组加减速的控制参数*)

	byParamIndex_Huang			: BYTE;
	uiControllerVel_Huang		: UINT;
	byFilmType					: BYTE;
	rFinalVel_ThisTime			: REAL;

	abyReserved					: ARRAY [1..28] OF BYTE;(*预留28个字节*)

	astTaperPoint_Rw						: ARRAY [1..10] OF StPoint_XY;
	(*新增工艺参数|2025.08.15.152008*)
	byFreqUpper_ExhaustAir :BYTE;
	uiFreqCoeff_Auto_ExhaustAir:UINT;
	byFreqMax_ExhaustAir:BYTE;
	byFreqMin_ExhaustAir:BYTE;

(*2025.8.19.205954*)
	xWorkMode_ManuAdj: BOOL;
	(*新增等料长相关参数|wang.nt|2025.08.20.220737*)
	lrFilmLen_UnwindToPU1					: LREAL;(*放料裁切点到1U的料膜距离|单位:mm|*)
	lrFilmLen_NotAdjFront					: LREAL;(*裁切点前不调整的料长|单位:mm|*)
	lrFilmLen_NotAdjBack					: LREAL;(*裁切点后不调整的料长|单位:mm|*)
	(*预套准相关变量|wang.nt|2025.08.21.162056*)
	byTurnOverAxisId						: BYTE;(*翻料架轴id@比如第10色反印那么 byTurnOverAxisId=10*)
	xPreRegisterAxisId_Manu					: BOOL;(*预套准的轴号手动确定@不考虑联动开关*)
	xSwitch_TempFromEnc_PT1000_If							: BIT;
	xSwitch_MotorTemp_PT1000_NTC_If						: BIT;
	xSwitch_TempFromEnc_PT1000_Of							: BIT;
	xSwitch_MotorTemp_PT1000_NTC_Of						: BIT;
//增加预热风和预加热参数2025.10.15.162208|niuj||88-16=72
	rHz_PreHotAir_ManuallySet							: REAL;(*预热风频率*)
	rSV_PreHeating										: REAL;(*预加热温控SV*)
	rCoeff_Scraper_Auto									: real;(*主刮刀自动系数*)

END_STRUCT
END_TYPE

{IMPLEMENTATION}

(* ---- StSysParam_Save.st ---- *)
(*@CES
Name=StSysParam_Save
Type=Gvl
TypeGuid=2db5746d-d284-4425-9f7f-2663a34b0ebc
Guid=a67fb49f-2618-48db-a2b1-8f99cf5bed12
HasDeclaration=True
HasImplementation=False
*)
{DECLARATION}
{attribute 'pack_mode' := '1'}
TYPE StSysParam_Save :
STRUCT
	dwFileVersion								: DWORD;(* 文件版本/后续作为识别参数的规范 *)
	iCustomerId									: INT;(* 客户id/2021.11.21.191558 *)
	dwEquipmentProf								: DWORD;(* 设备描述标志 *)
												(*bit0:反手机
												bit1:卫星式柔印
												bit2:机组式柔印

												bit3:凹印
												bit4:胶印
												bit5:品字形柔印
												bit8:特殊厂家显示界面-根据ID设置了

												bit20：双收双放
												bit21：A放B收
												bit22：收放料伺服控制

*)
	iUnitMaxNum									: INT;(* 最大色组数量 *)
	iCurveViewMaxRange				:INT;(*误差曲线量程上限		*)
	iUid							: INT;(*当前采样操作色组号*)

	(* 有关HMI字体高度设定的 *)
	iTitleTextHeight							: INT:=16;(* 标题字体高度 *)
	iEntryTextHeight							: INT:=12;(* 输入框字体高度 *)
	iLabelTextHeight							: INT:=12;(* 标签字体高度 *)
	iButtonTextHeight							: INT:=10;(* 按钮字体高度 *)
	iMessageTextHeight							: INT:=18;(* 消息字体高度 *)
	iRsvdTextHeight								: INT;(* 保留的字体高度 *)
	byLanguageId								: BYTE;(* 系统操作语言 *)
	byMinutes_ScrSaver							: BYTE;(* 屏幕延时分钟数 *)
	iPointDensity_RS							: INT;
	wCtlFlag_IndependentSettings				: WORD;
		(* 独立设定参数的标志
		/bit0=1底辊周长独立设置
		/bit1=1版辊周长独立设置
		/bit2=1网辊周长独立设置
		/bit3=1张带辊周长独立设置(保留)
		/bit4=1版辊压力电机丝杆节距独立设置
		/bit5=1版辊压力电机减速比独立设置
		/bit6=1网辊压力电机丝杆节距独立设置
		/bit7=1网辊压力电机减速比独立设置
		/bit8=1底辊减速比独立设置
		/bit9=1版辊减速比独立设置
		/bit10=1网辊减速比独立设置
		/bit11~bit15(保留)
		/ *)
(*原dwControlComplexBits内容不再用，直接拆分为BIT类型，直接不用*)

	xFlag_CancelSafetyGrate						: BIT;(*原dwControlComplexBits.14|取消光栅保护*)
	xSwitch_ArcTest_V							: BIT;(*原dwControlComplexBits.11|纵向快调标志*)
	xSwitch_ArcTest_H							: BIT;(*原dwControlComplexBits.15|横向快调标志*)
	xAllowLinkageChangeInRunning				: BIT;(*bit.24: 伺服电机支持开机状态下的单联动切换*)
	xChangLinkageStsWhenPrint					: bit;(*bit18:印刷状态下可以切换单联动*)
(*	dwControlComplexBits						: DWORD;(* 整机控制位 *)*)
			(*	/以下的整理来自2020.10.15.161719|后续版本严格按照该分配来执行 *)
			(*	/.0 : 置位表示关闭日志存储功能(默认为FALSE) *)
			(*	/.1 : 置位表示整机运动按照电机额定转速中的下限值进行限速(默认TRUE) *)
			(*	/.2 : 置位要求印刷机显示冷风机图标 *)
			(*	/.3 : 置位要求隐藏误差历史曲线的报警数值 *)
			(*	/.4 : 置位要求隐藏误差历史曲线的误差数值 *)
			(*	/.5 : 置位要求隐藏印刷机中的电机温度显示 *)
			(*	/.6 : 置位要求印刷机显示热风机图标 *)
			(*	/.7 : 置位要求界面的综合误差修正能通过界面手动控制横向电机 *)
			(*	/.8 : 置位放料卷径估计使能标志 *)
			(*	/.9 : 置位收料卷径估计使能标志 *)
			(*	/.10: 置位放料裁切窄方波+微分量补偿使能标志 *)
			(*	/.11~13: 保留/2021.12.11.194448/hdp *)
			(*	/.14: 关闭预套准修正量自动计算功能(TRUE=关闭;FALSE=打开自动计算<默认值>)/2021.12.11.194401/hdp修正.bit10重复 *)
			(*	/.15: 置位套色快调使能开关/2021.12.11.194420/hdp修正.bit11重复 *)
			(*	/.16: 界面套色修正步进量0.05(TRUE)/0.01(FALSE)选择/2021.11.4.172153 *)
			(*	/.17: 反复切换状态用于表示触发清除历史误差曲线的请求/2021.11.4.172150 *)
			(*	/.18: 套色报警使能开关/2021.11.4.180006 *)
			(*	/.19: Modbus通讯使能 *)
			(*	/.20: 横向采用步进控制 *)
			(*	/.22: 断料保护功能位 *)
			(*	/.26: 要求从站可以在空转状态下输入距离来进行纵向的快速对版 *)
			(*	/.29: 放料变频自调整使能(TRUE表示自调整) *)
			(*	/.30: DLL的粗采样波形显示采用形式(TRUE=方波;FALSE=模拟)
				/.31: 下伺服开关  *)
	astStMechanicalParamBuf						: ARRAY [1..5] OF StMechanicalParamBuf;(*2019.4.8.152905|新增系统机械参数|*)
	dwCtlSwitchRef						: DWORD;//整机控制位
													//.0: 伺服电机支持开机状态下的单联动切换
													//.1：色组联动采用按钮/开关
													//.2: 同步带长使用平均，True是平均，false是跟某一色
													//.3: 系统张力调整开关

//	byHorz_CtrlMode: BYTE;(*横向电机控制方式：0-不控制；1-同步电机；2-步进电机；3-伺服电机；--待续*)
	byRsvdata0							: BYTE;(*2025.9.16.093903*)
	rStepDrivePosPPulse					: REAL;(*步进电机|每个脉冲对应的位置值 mm|default.0.0002||*)
	iStepDrivePulsePRev					: INT;(*步进电机|每一圈对应的脉冲数|default.6000||*)
	iStepDriveSa_Vel					: INT;(*步进电机|步进电机启动速度,不能写0|default.10||*)
	iStepDrivePreReg_Vel				: INT;(*步进电机|步进电机预套准速度|default.50||*)
	iStepDriveManu_Vel					: INT;(*步进电机|步进电机手动调整低速速度|default.20||*)
	iStepDriveAuto_Vel					: INT;(*步进电机|步进电机自动调整速度|default.20||*)
	iStepDriveAccTime					: INT;(*步进电机|步进电机升速时间ms|default.50||*)
	iStepDriveManu_Vel_Fast				: INT;(*步进电机|步进电机手动高速调整速度|default.40||*)
	byOverPercent_RatedRpm				: BYTE;(*2019.4.17.163614|超频比例|相对于电机额定转速|*)
	rCurrent_Limit						: REAL;
	xWorkMode_Inch						: BOOL;(*单运行模式-TURE:按一下走一下听*)
(* 2021.2.4.141533 增加横向控制时的参数|34 bytes/lyt *)
	rHorCtl_PosPPulse					: REAL; (* 横向伺服控制每个脉冲对应的位置值 um|default.0.635| *)
	diHorCtl_PulsePRev					: DINT; (* 伺服电机脉冲/圈|default.131072 *)
	rHorCtl_PreReg_Vel					: REAL; (* 伺服电机预套准速度mm/sdefault.2 *)
	rHorCtl_Manu_Vel					: REAL; (* 伺服电机手动低速度mm/sdefault.0.5 *)
	rHorCtl_Manu_Vel_Fast				: REAL; (* 伺服电机手动高速度mm/sdefault.1 *)
	rHorCtl_Auto_Vel					: REAL; (* 伺服电机自动速度mm/sdefault.0.5 *)
	iHorCtl_Num							: INT; (* 横向控制电机侧|default.60 *)
	iHorCtl_Den							: INT; (* 横向控制传动侧|default.1 *)
	rHorCtl_Pitch						: REAL; (* 横向控制螺距mm|default.5 *)
	iHorCtl_AccDecTime					: INT; (* 加速到自动速度或者自动速度减速到0的时间ms|default.10 *)
	(*2023.8.29.151955增加报警铃响铃时间*)
	diTimeHold_Prestart				:DINT;
	diTimeHold_Uw_Diam				:DINT;
	diTimeHold_Rw_Diam				:DINT;
	diTimeHold_Rw_Prnlength			:DINT;

	byHotBlowerStopDelayTime					: BYTE;//热风延时关闭时间
	byHeatingOutWay_III							: BYTE;
	iTimeOut_Slave_485_Inverter				: INT;

(*2023.3.27.151009需增加排风、递墨、热风、刮刀485控制使能开关-用于屏蔽相关报警||
新增水加热控制系数-分段*)

	iCofe_TempCtl_30						: INT;(*温度偏差超过30℃-系数-水加热推荐30，蒸汽加热推荐50*)
	iCofe_TempCtl_30_10						: INT;(*温度偏差超过30℃-10℃-系数-水加热推荐40，蒸汽加热推荐100*)
	iCofe_TempCtl_10_5						: INT;(*温度偏差超过10℃-5℃-系数-水加热推荐50，蒸汽加热推荐100*)
	iCofe_TempCtl_5							: INT;(*温度偏差5℃以内-系数-水加热推荐60，蒸汽加热推荐100*)
	iTime_Thres_Water						: INT;(*水加热/蒸汽加热阀门打开时间-用于计算最大调整量*)
	byHeatingMode							: BYTE;(*0:加热模块1：驱动器温控2：温控表*)

	byOverTempValue						: BYTE;(* 2022.3.21.184802/过温值/摄氏度 *)

	byEn_ExtraFun_485						: BYTE;
	iPidAlgorithm_Threshold					: INT;(*PID;(*pid算法介入阈值(相差一定温度后进入pid算法调整)|目标速度-当前速度>该值-*) *)
	iMaxOutValue								: INT;(*最大输出值|长有效的最大值*)
	rKp											: REAL;(*i_rKp:REAL;(*Kp*)      *)
	rKi											: REAL;(*i_rKi:REAL;(*Ki*)    *)
	rKd											: REAL;(*i_rKd:REAL;(*Kd*)    *)
	uiCtrolCycle_Ms							: UINT;(*i_uiCtrolCycle_Ms:UINT;(*控制周期|ms*)   *)
(*2022.10.22.131113*)

(*iWaterValue_Threshold|2022.10.27.184352|水加热阀值*)
	iWaterValue_Threshold					: INT;
	iTempAcc_Threshold						: INT;(*温度上升速率阀值*)
	iDecSV_PV_Threshold					: INT;(*温度阀值2022.10.28.155136*)
	(*2023.12.21.210222||xi.hy||停机后关闭加热使能/停机后关闭热风使能/热风延时关闭时间*)
	xEn_HeatOff_AfterStop:BOOL;
	xEn_HeatAirOff_AfterStop:BOOL;
	rDelayOff_HotAir:REAL;
	(*2024.06.11.102646*)
	iDebugStep								: INT	:=0;(*初始值0||调试向导|2018.12.19.134002||*)
	dwSwitch								: DWORD	:=0;(*初始值0||调试向导|2018.12.19.134002||*)
												(*标志位使用介绍：
												* 控制调试界面确认完成标志
												* bit.0: 调试向导DEBUGSTEP_CONFIG系统配置界面完成标志|
												* bit.1: 调试向导DEBUGSTEP_FUNCTIONSET功能配置完成标志|
												* bit.2: 调试向导DEBUGSTEP_CHECKPARAM1核对参数1完成标志|
												* bit.3: 调试向导DEBUGSTEP_CHECKPARAM2核对参数2完成标志|
												* bit.4: 调试向导DEBUGSTEP_CHECKPARAM3核对参数3完成标志|
												* bit.5: 调试向导DEBUGSTEP_AXISIO色组IO测试完成标志|
												* bit.6: 调试向导DEBUGSTEP_UWRWIO收放料IO测试完成标志|
												* bit.7: 调试向导DEBUGSTEP_ANALOGIO模拟量测试完成标志|
												* bit.8: 调试向导DEBUGSTEP_EXTRAPARAM扩展参数完成|
												|*)
//2026.5.8.160853调整强度切换标志

//2026.4.25.144455增加调整强度切换开关变量|1个字节|2-1=1
	byArcIntensity								: BYTE;
//2026.4.25.144533
	byData:								 BYTE;(*原纵横向飞点阈值*)

	uiMaxVel_UseCalcAcc				: UINT;
	xUnitPressOneBtn			: BOOL := FALSE; (* 色组合压离压单个按钮标志 *)
	xAllPressOneBtn				: BOOL := FALSE; (* 全体合压离压单个按钮标志 *)
	xPreCutOneBtn_Uw			: BOOL := FALSE; (* 接料准备解除单个按钮标志_放料 *)
	xPreCutOneBtn_Rw			: BOOL := FALSE; (* 接料准备解除单个按钮标志_收料 *)

	xTypeGetInitDiam						: BOOL;(*方式切换|TRUE=使用停机之前的值|=FALSE 使用固定值*)
	uiMaxDia								: UINT;(*最大的卷径@mm*)
	uiInitDiam_Uw							: UINT;(*初始的卷径@mm|=0 按照200---uiMaxDia取中间值*)
	uiInitDiam_Rw							: UINT;(*初始的卷径@mm|=0 按照200---uiMaxDia取中间值*)
	xAutoSetArcCtlWay						: BOOL;(*自动设置耦合方式@根据是否隔色控制*)
	byCouplingType:BYTE:=0;(*耦合方式@=0原来的直接传递的逻辑@不输出耦合量
									 @=1新修改的按照比例定位传递。总量100%@从o_aiCouplingValue_A输出
									 @=2新修改的按照比例定位传递。总量根据输入的耦合值@从o_aiCouplingValue_A输出
									 @=3调整引起张力变化需要直接传递一定比例-等到达下一色取消这部分传递o_aiCouplingValue_T输出、
									   等待固定料长传递之前调整的量o_aiCouplingValue_A输出*)
(*新增加参数|wang.nt|2025.08.07.143540*)
	wMachineArchitectureRef : WORD;(*机器架构描述*)
	iPromptMsgId : INT;(*提示信息ID（报警代码）*)
	byHorzCtlMode : BYTE;(*横向控制方式-同步-步进-伺服*)
	byCheckTimeToTips_BrakeResistance : BYTE;(*制动电阻访问超限提示时间*)
	byCheckTimeToEStop_BrakeResistance : BYTE;(*制动电阻访问超限急停时间*)
	byAccessTimes_BrakeResistance : BYTE;(*制动电阻报警限制*)
	byAlarmHold_VOL_Uw : BYTE;(*放料没料响应时间*)
	byAlarmHold_PrnLength :BYTE;(*收料印长报警响应时间*)
	rOpenThr_Ele : REAL;(*电加热开启*)
	rCloseThr_Ele : REAL;(*电加热关闭*)
	rDealValue_Water : REAL;(*水加热死区*)
	iHeatingDebugValue_Water : INT;(*测试开度*)
	diStepDriveDebugPulse : DINT;(*测试脉冲数*)
	rStepDriveDebugPulse_PosAct :REAL;(*测试距离*)
	iStepDriveDebugNum : INT;(*测试色组号*)
	rHz_MainExhaust_ManuallySet : REAL;(*主排风设定频率*)
	byFreq_I_ExhaustAir : BYTE;(*排风一档频率*)
	byFreq_II_ExhaustAir : BYTE;(*排风二档频率*)
	byFreq_III_ExhaustAir : BYTE;(*排风三档频率*)
	(*9905界面参数*)
	byPseudoRandomRoundTimes:BYTE;
	rPseudoRandomAmplitude:REAL;
	bySetTestPid_IfOf:BYTE;
	by10vSignalCoef:BYTE;
	rCompensateGirthWhenAccing_If	:REAL;
	rCompensateGirthWhenAccing_Of	:REAL;
	byArcDeCoupleStepTest			:BYTE;
	iCustomerLogoOffsetX			:INT;
	byGuardrialColor_R				:BYTE;
	byGuardrialColor_G				:BYTE;
	byGuardrialColor_B				:BYTE;
	iLedFuncId						:INT;
	iSetHmiResValue					:INT;
	wRunningTime_Day				:WORD;
	byRunningTime_Hour				:BYTE;
	byRunningTime_Min				:BYTE;
	byRunningTime_Sec				:BYTE;
	byArcIntensity_W				:BYTE;
	byArcIntensity_M				:BYTE;
	byArcIntensity_S				:BYTE;
	byMotorOverTempValue_UseEncTemp	:BYTE;
	byRemainSpaceNum_PTCTL			:BYTE;
	rSpeed_SCoeff_Type789			:REAL;
	byMaxPulseOut_16dIO				:BYTE;
	bySysSamplePrecision			:BYTE;
	byArcAdjValueDealType			:BYTE;
	byArcErrLimitToCtl_P			:BYTE;
	byArcErrLimitToCtl_I 			:BYTE;
	byMaxPulseOut_Module			:BYTE;
	byArcFineSampleType				:BYTE;
	byArcPidGetType 				:BYTE;
	rFilmLenth_Eyes					:REAL;
	uiArcSysDelayTime_ms           	:UINT;
	byParamIndex_Huang				:BYTE;
	uiControllerVel_Huang			:UINT;
	byDeCoupleArcNum				:BYTE;

(*部分开关-直接用BIT-先放这里2025.8.8.151629*)
	xSwitch_PreHotEn_Print					 :BIT;(*预热印刷激活开关*)
    xSwitch_ExhAir_Limit_HotWind			 :BIT;(*排风限制热风开关*)
    xSwitch_ExhAir_Limit_Run				 :BIT;(*排风限制开机开关*)
    xSwitch_CommEn_WatchDevice_Tcp			 :BIT;(*TCP-外部监控设备开关*)
    xSwitch_CommEn_WatchDevice_485			 :BIT;(*485-外部监控设备开关*)
    xSwitch_CommEn_1U_485					 :BIT;(*1色人机通讯开关*)
    xSwitch_CommEn_485						 :BIT;(*485通讯开关*)
    xSwitch_CommEn_485_Exh					 :BIT;(*排风485通讯开关*)
    xSwitch_CommEn_485_Scraper				 :BIT;(*刮刀485通讯开关*)
    xSwitch_CommEn_485_InkRoller			 :BIT;(*递墨辊485通讯开关*)
    xSwitch_CommEn_485_HotWind				 :BIT;(*热风485通讯开关*)
    xSwitch_ArcIntensityBtn_Hmi				 :BIT;(*手动调节随速度走开关*)
    xSwitch_PrnRatioIndividual_Setting		 :BIT;(*色组版辊减速比单独设置开关*)
    xSwitch_NetRatioIndividual_Setting		 :BIT;(*色组网辊减速比单独设置开关*)
    xSwitch_BottomRatioIndividual_Setting	 :BIT;(*色组底辊减速比单独设置开关*)
    xSwitch_StepDriveDebugRun				 :BIT;(*横向步进电机测试执行开关*)

	xSetProPointEn										: BIT;
	xUseMaxTimeAsSBegin_InLowSpeed      				: BIT;
	xPseudoRandomEn                     				: BIT;
	xPseudoRandomStart                  				: BIT;
	xEn_RevLimit                        				: BIT;
	xSaveFineSampleData_ToArc           				: BIT;
	xReqSetLedFunc                      				: BIT;
	xSetHmiResolution                   				: BIT;
	xPopupWindowVisible                 				: BIT;
	xInitArcErr_AjdImmediately          				: BIT;
	xPhaseAutoRecoveryEn                				: BIT;
	xKeepServo_PreRegisterDne           				: BIT;
	xUseIfVel_Uw                        				: BIT;
	xKeepServo_Stop                     				: BIT;
	xAxisPrfVelEn                       				: BIT;
	xUseGc_PID_2025                     				: BIT;
	xFlag_Follow_1U_Double_V            				: BIT;
	xArcErrCorrectIsRev_V               				: BIT;
	xAutoSetSampleType                  				: BIT;
	xGetSampleTypeBtn                   				: BIT;
	byKadj_SetType				: BYTE;
	xUseArcErr_Lp				: BOOL;(*套色误差使用低通*)
	byUseArcAccOrDecCompensate	: BYTE;

	(*新增参数-开始|wang.nt|2025.08.12.141656*)
	byAlarmHold_CutDne_Uw		: BYTE := 3; (* 放料接完料后报警持续时间@单位s *)
	(*新增参数-结束|wang.nt|2025.08.12.141656*)
	(*新增工艺参数|2025.08.15.152053*)
	iDelayMsec_HeatBlower :INT ;//热风停止延时
	xAirExhaustLimit:BOOL;(*排风限制开机*)
	(*2025.8.19.211236*)
	byTypeFollow_Arc	: BYTE;

	iRemaindPartCouplingPos	: INT:=0;(*剩余部分的耦合位置@距离总幅数
														   @=1 到达下一色前第一幅
														   @=2 到达下一色前第二幅*)
	(*新增等料长参数|wang.nt|2025.08.20.221817*)
	dwAxis_SkipTheHeader				: DWORD;(*让料头标志| 位标志bit0=机组1,...,bit31=机组32*)
	(*新增预套准参数|2025.08.23.091002*)
	byMechanicalTypeId					: BYTE;(*1摆臂\2直压\3pvc直压|*)
	xFilpSwitch:BOOL;(*翻转架开关*)
(*全局*)
(*要更新数据结构2025.10.13.134149--这些全部要加到金刚读写通讯区域*)
	(*2025.6.9.142100+油墨槽控制@20BYTES*)
	xInkGrooveCtlEn						: BOOL;(*油墨槽控制使能*)
	xInkGrooveCtlDirRev					: BOOL;(*油墨槽运动方向取反*)
	iInkGroovePulsePRev					: INT;(*一圈的脉冲数*)
	iInkGrooveSa_Vel					: INT;(*油墨槽控制|油墨槽控制启动速度,不能写0|default.10||*)
	iInkGroove_Vel						: INT;(*油墨槽控制|油墨槽控制手动调整速度|default.20||*)
	iInkGrooveAccTime					: INT;(*油墨槽控制|油墨槽控制升速时间ms|default.50||*)
	rInkGroovePosPPulse					: REAL;(*油墨槽控制|每个脉冲对应的位置值 mm|default.0.0002||*)
	iInkGrooveMoveDis_Max				: INT;(*油墨槽控制|最大运行的距离 mm|*)

	(*增加排风三档频率|2022.5.5.154339*)
	(*增加了热风三档频率|2022.5.6.083338*)
	byFreq_I_AirHot						: BYTE;
	byFreq_II_AirHot					: BYTE;
	byFreq_III_AirHot					: BYTE;
//2025.10.20.145004增加排风控制相关一些变量72-5=67
	byExhaustMode				: BYTE;
	byExhaustLinkageNum			: BYTE;
	byFreqMax_ExhaustAir		: BYTE;
	byFreqMin_ExhaustAir		: BYTE;
	byCoefExhaust				: BYTE;
	xArcFollowAnyAxis			: BOOL;
	byTypeFollow1UEn			: BYTE;
	xFlag_Follow_1U_Double_H	: BOOL;
	byModbusNum_Max							: BYTE;

END_STRUCT
END_TYPE

{IMPLEMENTATION}

(* ---- StUnitParam_Save.st ---- *)
(*@CES
Name=StUnitParam_Save
Type=Gvl
TypeGuid=2db5746d-d284-4425-9f7f-2663a34b0ebc
Guid=eeacd55f-9111-4e09-ad6b-b078dffd0b62
HasDeclaration=True
HasImplementation=False
*)
{DECLARATION}
{attribute 'pack_mode' := '1'}
TYPE StUnitParam_Save :
STRUCT
	byGrpId										: BYTE;(*系ID*)
	rGirth_BottomRoller							: REAL;(* 底辊周长 *)
	uiNum_BottomRoller							: UINT;(* 底辊减速比分子 *)
	uiDen_BottomRoller							: UINT;(* 底辊减速比分母 *)
	rGirth_PrnRoller							: REAL;(* 版辊周长 *)
	uiNum_PrnRoller								: UINT;(* 版辊减速比分子 *)
	uiDen_PrnRoller								: UINT;(* 版辊减速比分母 *)
	rGirth_NetRoller							: REAL;(* 网辊周长 *)
	uiNum_NetRoller								: UINT;(* 网辊减速比分子 *)
	uiDen_NetRoller								: UINT;(* 网辊减速比分母 *)
	rLength_Band								: REAL;(* 带长 *)
	rErrLength_Band								: REAL;(* 设置带长与实际检测之间的误差 *)
	rGirth_StrRoller							: REAL;(* 张带辊周长 *)
	uiNum_StrRoller								: UINT;(* 张带辊减速比分子 *)
	uiDen_StrRoller								: UINT;(* 张带辊减速比分母 *)
	rScrewPitch_Horz							: REAL;(* 横向架丝杆节距/整机设置状态/单位mm *)
	uiNum_Horz									: UINT;(* 横向电机减速比分子/整机设置状态 *)
	uiDen_Horz									: UINT;(* 横向电机减速比分母/整机设置状态 *)
	lrLimit_Operate_Horz						: LREAL;(*操作侧电机限位*)
	lrLimit_Driver_Horz							: LREAL;(*传动侧电机限位*)
	wCtlmod_PrnRoller_Pressure					: WORD;(* 版辊压力控制方式 *)
		(*
		/0表示不控制(默认)
		/1为独立单轴控制
		/2为双轴控制
		/4为4轴驱动器控制 *)
	rScrewPitch_PrnRoller_Pressure				: REAL;(* 版辊压力架丝杆节距/单位mm *)
	uiNum_PrnRoller_Pressure					: UINT;(* 版辊压力电机减速比分子 *)
	uiDen_PrnRoller_Pressure					: UINT;(* 版辊压力电机减速比分母 *)
	rScrewPitch_NetRoller_Pressure				: REAL;(* 网辊压力架丝杆节距/单位mm *)
	uiNum_NetRoller_Pressure					: UINT;(* 网辊压力电机减速比分子 *)
	uiDen_NetRoller_Pressure					: UINT;(* 网辊压力电机减速比分母 *)
	rScrewPitch_StrRoller_Pressure				: REAL;(* 张带辊压力架丝杆节距/单位mm *)
	uiNum_StrRoller_Pressure					: UINT;(* 张带辊压力电机减速比分子 *)
	uiDen_StrRoller_Pressure					: UINT;(* 张带辊压力电机减速比分母 *)
	rMovementHiSpd_PrnRoller_Pressure			: REAL;(* 版辊压力架移动速度(高)/默认单位:mm/s *)
	rMovementHiSpd_NetRoller_Pressure			: REAL;(* 网辊压力架移动速度(高)/默认单位:mm/s *)
	rMovementLoSpd_PrnRoller_Pressure			: REAL;(* 版辊压力架移动速度(低)/默认单位:mm/s *)
	rMovementLoSpd_NetRoller_Pressure			: REAL;(* 网辊压力架移动速度(低)/默认单位:mm/s *)
	rPos_press_dn_PrnRoller_Pressure_M			: LREAL;(* 合压位置/版辊压力电机M侧/单位:mm *)
	rPos_press_dn_PrnRoller_Pressure_G			: LREAL;(* 合压位置/版辊压力电机G侧/单位:mm *)
	rPos_press_up_PrnRoller_Pressure_M			: LREAL;(* 离压位置/版辊压力电机M侧/单位:mm/根据当前合压位置实时变化/2021.12.29.140151 *)
	rPos_press_up_PrnRoller_Pressure_G			: LREAL;(* 离压位置/版辊压力电机G侧/单位:mm/根据当前合压位置实时变化/2021.12.29.140151 *)
	rPos_load_unload_PrnRoller_Pressure_M		: LREAL;(* 装卸辊位置/版辊压力电机M侧/单位:mm *)
	rPos_load_unload_PrnRoller_Pressure_G		: LREAL;(* 装卸辊位置/版辊压力电机G侧/单位:mm *)
	rPos_press_dn_NetRoller_Pressure_M			: LREAL;(* 合压位置/网辊压力电机M侧/单位:mm *)
	rPos_press_dn_NetRoller_Pressure_G			: LREAL;(* 合压位置/网辊压力电机G侧/单位:mm *)
	rPos_press_up_NetRoller_Pressure_M			: LREAL;(* 离压位置/网辊压力电机M侧/单位:mm/根据当前合压位置实时变化/2021.12.29.140151 *)
	rPos_press_up_NetRoller_Pressure_G			: LREAL;(* 离压位置/网辊压力电机G侧/单位:mm/根据当前合压位置实时变化/2021.12.29.140151 *)
	rPos_load_unload_NetRoller_Pressure_M		: LREAL;(* 装卸辊位置/网辊压力电机M侧/单位:mm *)
	rPos_load_unload_NetRoller_Pressure_G		: LREAL;(* 装卸辊位置/网辊压力电机G侧/单位:mm *)
	rPos_press_dn_StrRoller_Pressure_M			: LREAL;(* 合压位置/网辊压力电机M侧/单位:mm *)
	rPos_press_dn_StrRoller_Pressure_G			: LREAL;(* 合压位置/网辊压力电机G侧/单位:mm *)
	rPos_press_up_StrRoller_Pressure_M			: LREAL;(* 离压位置/网辊压力电机M侧/单位:mm/根据当前合压位置实时变化/2021.12.29.140151 *)
	rPos_press_up_StrRoller_Pressure_G			: LREAL;(* 离压位置/网辊压力电机G侧/单位:mm/根据当前合压位置实时变化/2021.12.29.140151 *)
	rPos_load_unload_StrRoller_Pressure_M		: LREAL;(* 装卸辊位置/网辊压力电机M侧/单位:mm *)
	rPos_load_unload_StrRoller_Pressure_G		: LREAL;(* 装卸辊位置/网辊压力电机G侧/单位:mm *)
	rGirth_Confirmed_press_dn_PrnRoller			: REAL;(* 确认合压位时候的版辊周长*)
	rGirth_Confirmed_press_dn_NetRoller			: REAL;(* 确认合压位时候的网纹辊周长*)
	rGirth_Confirmed_press_dn_StrRoller			: REAL;(* 确认合压位时候的网纹辊周长*)

//2024.12.05.180655 | bai.zy | 下面两个BYTE类型的标志不用了，合成一个WORD标志，做一下压力相关功能的参数
///////////////////////////////////////////////////////////////////////////////////////////////////
(* 2021.12.25.083025/hdp/按照2021.12.24试机完成后lyt同步的工程进行注释更新 *)
// 	(*判定规划器和编码器的方向|*)
// 	(*FALSE-编码器方向和规划器方向一致|TRUE-编码器方向和规划器方向不一致*)
// 	bySts_PrfPosAndEncPosDir:BYTE;(*/.0 版辊操作侧压力电机方向
// 									/.1 版辊操作侧压力电机方向确认完成了
// 									/.2 版辊传动侧压力电机方向
// 									/.3 版辊传动侧压力电机方向确认完成了
// 									/.4 网纹辊传动侧压力电机方向
// 									/.5 网纹辊传动侧压力电机方向确认完成了
// 									/.6 网纹辊传动侧压力电机方向
// 									/.7 网纹辊传动侧压力电机方向确认完成了*)
//
// 	(*实际编码器方向|FALSE-实际编码器方向和规划器方向一致|TRUE-实际编码器方向和规划器方向不一致*)
// 	bySts_PrfPosAndActEncPosDirDir:BYTE;(*/.0 版辊操作侧压力电机方向
// 									/.1 版辊操作侧压力电机方向确认完成了
// 									/.2 版辊传动侧压力电机方向
// 									/.3 版辊传动侧压力电机方向确认完成了
// 									/.4 网纹辊传动侧压力电机方向
// 									/.5 网纹辊传动侧压力电机方向确认完成了
// 									/.6 网纹辊传动侧压力电机方向
// 									/.7 网纹辊传动侧压力电机方向确认完成了*)
// (* end/hdp *)
// (* end/hdp *)
////////////////////////////////////////////////////////////////////////////////////////////////////
	wFlag_PressFun		: WORD;(*.0: 色组安装手轮开关
									.1 版辊压力粗细调
									.2 网辊压力粗细调
									.3 张带压力粗细调*)

	lrAbsEncZeroPos_PrnRoller_Pressure_M		: LREAL;(* 版辊压力电机绝对值位置M侧/零位 *)
	lrAbsEncZeroPos_PrnRoller_Pressure_G		: LREAL;(* 版辊压力电机绝对值位置G侧/零位 *)
	lrAbsEncZeroPos_NetRoller_Pressure_M		: LREAL;(* 网辊压力电机绝对值位置M侧/零位 *)
	lrAbsEncZeroPos_NetRoller_Pressure_G		: LREAL;(* 网辊压力电机绝对值位置G侧/零位 *)

	lrAbsEncLimMin_PrnRoller_Pressure_M			: LREAL;(* 版辊压力电机绝对值位置M侧边界min *)
	lrAbsEncLimMax_PrnRoller_Pressure_G			: LREAL;(* 版辊压力电机绝对值位置G侧边界max *)
	lrAbsEncLimMin_NetRoller_Pressure_M			: LREAL;(* 网辊压力电机绝对值位置M侧边界min *)
	lrAbsEncLimMax_NetRoller_Pressure_G			: LREAL;(* 网辊压力电机绝对值位置G侧边界max *)
	xConfirmAbsEncZeroPosDne_PrnRoller_Pressure_M	: BOOL;(* 版辊压力电机绝对值位置M侧/零位确认完成 *)
	xConfirmAbsEncZeroPosDne_PrnRoller_Pressure_G	: BOOL;(* 版辊压力电机绝对值位置G侧/零位确认完成 *)
	xConfirmAbsEncZeroPosDne_NetRoller_Pressure_M	: BOOL;(* 网辊压力电机绝对值位置M侧/零位确认完成 *)
	xConfirmAbsEncZeroPosDne_NetRoller_Pressure_G	: BOOL;(* 网辊压力电机绝对值位置G侧/零位确认完成 *)

(* 2021.12.29.140315/hdp/lyt *)
	xConfirmload_unloadPosDne_PrnRoller_Pressure_M	: BOOL;(* 版辊压力电机换版位置M侧/确认完成 *)
	xConfirmload_unloadPosDne_PrnRoller_Pressure_G	: BOOL;(* 版辊压力电机换版位置G侧/确认完成 *)
	xConfirmload_unloadPosDne_NetRoller_Pressure_M	: BOOL;(* 网辊压力电机换版位置M侧/确认完成 *)
	xConfirmload_unloadPosDne_NetRoller_Pressure_G	: BOOL;(* 网辊压力电机换版位置G侧/确认完成 *)

	xConfirmDnPosDne_PrnRoller_Pressure_M			: BOOL;(* 版辊压力电机合压位置M侧/确认完成 *)
	xConfirmDnPosDne_PrnRoller_Pressure_G			: BOOL;(* 版辊压力电机合压位置G侧/确认完成 *)
	xConfirmDnPosDne_NetRoller_Pressure_M			: BOOL;(* 网辊压力电机合压位置M侧/确认完成 *)
	xConfirmDnPosDne_NetRoller_Pressure_G			: BOOL;(* 网辊压力电机合压位置G侧/确认完成 *)
	xEnable_arc									: BOOL;(* 套印使能标志 *)
	iMarkTypeId									: INT;(* 标记形式 *)
	iMarkArrangeMode							: INT;(* 标记排列方式 *)
	iGateWidthPhy								: INT;(* 波门宽度/单位:mm *)
	iGateWidthRoundPoints						: INT;(* 波门宽度占据的粗采样点数 *)
	iGateWidthFinePoints						: INT;(* 波门宽度占据的精采样点数 *)
	iGateSa										: INT;(* 波门地址1 *)
	iGateSaEx									: INT;(* 波门地址2 *)
	rAlr_V										: REAL;(* 纵向报警值/pdu通信协议采用x100整型传输 *)
	rAdj_V										: REAL;(* 纵向版修正 *)
	byAvg_V										: BYTE;(* 纵向平均值 *)

	iKp_V										: INT;(* 纵向Kp *)
	iKi_V										: INT;(* 纵向Ki *)
	iKd_V										: INT;(* 纵向Kd *)
	rDeadzoneMin_V								: REAL;(* 纵向不工作区/小/pdu通信协议采用x100整型传输 *)
	rAlr_H										: REAL;(* 横向报警值/pdu通信协议采用x100整型传输 *)
	rAdj_H										: REAL;(* 横向版修正 *)
	byAvg_H										: BYTE;(* 横向平均值 *)

	iKp_H										: INT;(* 横向Kp *)
	iKi_H										: INT;(* 横向Ki *)
	iKd_H										: INT;(* 横向Kd *)
	rDeadzoneMin_H								: REAL;(* 横向不工作区/小/pdu通信协议采用x100整型传输 *)
	rDeadzoneMax_H								: REAL;(* 横向不工作区/大/pdu通信协议采用x100整型传输 *)
	lrPreReg_Length_V						: LREAL;(*纵向预套准料长值|单位:mm|*)
	lrFilmLengthFromPrevUnit				: LREAL;(*存储前色到当前色的压印点间料长|*)
	lrPreReg_Adjust							: LREAL;(*预套准调整量|*)
	dwFlag_Ctl									: DWORD;(* 控制标志 *)
(*												/bit0.横向开关 *)
(*												/bit1.门内基线 *)
(*												/bit2.T1反极性 *)
(*						dwFlag_Ctl						/bit3.T2反极性 *)
(*												/bit4.纵向调整反 *)
(*												/bit5.横向调整反 *)
(*												/bit6.双波门 *)
(*												/bit7.单标记调整反 *)
(*												/bit8.反印开关*)
(*												/bit9.电眼型号KSC012(A) *)
(*												/bit10.波门锁定 *)
(*												/bit11.T1反极性-第二个门内 *)
(*												/bit12.T2反极性-第二个门内 *)
(*												/bit13.T1小信号 *)
(*												/bit14.T2小信号 *)
(*												/ *)

(*												/bit28.套色方式-曜光/光电眼TRUE为曜光 *)
(*												/bit29.压力电机步进快慢选择/TRUE表示快挡位/2021.12.22.165105/hdp *)
(*												/bit30.KSC-012(A)光电眼两路DO设置-DO0 *)
(*												/bit31.KSC-012(A)光电眼两路DO设置-DO1 *)
(*												/ *)
	dwFlag_Sts									: DWORD;(* 状态标志 *)
(*												/bit0.纵向自动 *)
(*												/bit1.横向自动 *)
(*												/ *)
(*												/bit8.纵向跟任意色 *)
(*												/bit9.横向跟任意色 *)
(*												/bit12.纵向使用跟踪第一色色标计算误差-反之使用前一色色标计算|2023.09.14.102543 *)
(*												/bit13.横向使用跟踪第一色色标计算误差-反之使用前一色色标计算2023.09.14.102543 *)
(*												bit14=1  纵向使用间接跟1色误差反之-默认使用前一色
												bit15=1  横向使用间接跟1色误差-

												//bit30+bit31用作精采样数据滤波方式选择||2025.11.15.132316
												//00：均值滤波/01：低通滤波

*)
	diPreReg_AdjustVal_H					: DINT;(*预套准修正值-横向|单位:mm|*)
	lrAI_med_CoatingPrn						: LREAL;(*涂布中位值|*)
	xSwitchOn_CoatingPrn					: BOOL;(*涂布开关|*)
	xReverseAdj_CoatingPrn					: BOOL;(*涂布反向调整|*)
	byAdjMode_CoatingPrn					: BYTE;(*涂布调整方式|0~1|*)
	iKp_CoatingPrn							: INT;(*涂布Kp|0~500|*)
	iKi_CoatingPrn							: INT;(*涂布Ki|0~500|*)
	iKd_CoatingPrn							: INT;(*涂布Kd|0~500|*)
	bySensorType_CoatingPrn					: BYTE;(*涂布传感器类型|0~10|*)
	lrAI_CoatingPrn							: LREAL;(*涂布模拟量|*)
	lrGirth_Using_CoatingPrn				: LREAL;(*使用的涂布版周长|*)
	bySignalGain								: BYTE;(* 信号增益控制/2021.10.21.103435 *)
(*												/bit0~bit3.T1的信号增益 *)
(*												/bit4~bit7.T2的信号增益 *)
	xLinkage									: BOOL;(*色组联动*)
	rInversedPrecision						: REAL;(*系统精度2023.6.7.170657*)
	byCouplingMask							: BYTE;(*耦合开关|
													*.bit0=1: 纵向调整量传递|
													*.bit1=1: 横向调整量传递|
													*.bit2=1: 纵向误差传递|
													*.bit3=1: 横向误差传递|
													|*)
	rHigh_Prn_Roller					:REAL;//轴高
	rHigh_Net_Roller					:REAL;//轴高

	rweigth_Prn_Bottom_Confirm					: REAL;//标定位置时这个是版辊中心到版辊和底辊/中心辊切点的横向距离
	rweigth_Prn_Net_Confirm					: REAL;//标定位置时这个是版辊中心到版辊和网辊切点的横向距离
	rweigth_Net_Prn_Confirm					: REAL;//标定位置时这个是版辊中心到版辊和底辊/中心辊切点的横向距离
	rweigth_Net_Load_Confirm					: REAL;//标定位置时这个是版辊中心到版辊和网辊切点的横向距离

	dwColor_Print							: DWORD;//16进制颜色变量
													//16#FFFFFFFF分别代表
													//bit31-bit24:透明度
													//bit23-bit16:RED红色
													//bit15-bit8:GREEN绿色
													//bit7-bit0:BLUE蓝色
	wLines_Net_Roller						: WORD;//网纹辊线数
	rStep_Pressure_Prn_Net					: REAL;
	//2023.12.22.211317}||新增版辊网辊步进1928-1924
//bai.zy | 2024.01.15.105100 | 增加张带合压位换版位标定完成标志------2字节
	xConfirmDnPosDne_StrRoller_Pressure_M			: BOOL;(* 张带辊压力电机合压位置M侧/确认完成 *)
	xConfirmDnPosDne_StrRoller_Pressure_G			: BOOL;(* 张带辊压力电机合压位置G侧/确认完成 *)
//bai.zy | 2024.03.21.130939 | 增加印刷位,32字节
	lrEncPosPrintDn_Prn_M : LREAL;
	lrEncPosPrintDn_Prn_G : LREAL;
	lrEncPosPrintDn_Net_M : LREAL;
	lrEncPosPrintDn_Net_G : LREAL;
	lrEncPosPrintDn_Str_M : LREAL;
	lrEncPosPrintDn_Str_G : LREAL;

//2024.10.21.114530 | bai.zy | 版辊网辊操作侧传动侧平行位置标定值	48字节
	lrEncPosParallel_Prn_M : LREAL;
	lrEncPosParallel_Prn_G : LREAL;
	lrEncPosParallel_Net_M : LREAL;
	lrEncPosParallel_Net_G : LREAL;
	lrEncPosParallel_Str_M : LREAL;
	lrEncPosParallel_Str_G : LREAL;
//2024.10.21.114530 | bai.zy | 版辊网辊操作侧传动侧合压位偏移量	  48字节
	lrPrintPosOffsetDn_Prn_M : LREAL;
	lrPrintPosOffsetDn_Prn_G : LREAL;
	lrPrintPosOffsetDn_Net_M : LREAL;
	lrPrintPosOffsetDn_Net_G : LREAL;
	lrPrintPosOffsetDn_Str_M : LREAL;
	lrPrintPosOffsetDn_Str_G : LREAL;

//2024.10.22.180832||增加	adiEncPos_Start_Virtual_0				: ARRAY [1..MAX_UNIT_NUM] OF DINT; 4字节
	diEncPos_Start_Virtual_0: DINT;
//2024.11.26.125320 | 增加采样减速比		8字节
	diSampleNum : DINT;//采样减速比分子
	diSampleDen : DINT;//采样减速比分母

//2024.11.27.154753 | bai.zy | 增加绝对编码器位置,48字节
	liABSPos_Prn_M : LINT;
	liABSPos_Prn_G : LINT;
	liABSPos_Net_M : LINT;
	liABSPos_Net_G : LINT;
	liABSPos_Str_M : LINT;
	liABSPos_Str_G : LINT;
//2024.12.03.162342 | 增加调试阶段的压力运动	要大幅度运行必须平行 使用平行位置当做最小值  是否合理？？先用吧  --54字节
	axPressLimit_Min : ARRAY[1..3] OF BOOL;
	axPressLimit_Max : ARRAY[1..3] OF BOOL;

	lrEncPosLimit_Prn_M_Max : LREAL;
	lrEncPosLimit_Prn_G_Max : LREAL;
	lrEncPosLimit_Net_M_Max : LREAL;
	lrEncPosLimit_Net_G_Max : LREAL;
	lrEncPosLimit_Str_M_Max : LREAL;
	lrEncPosLimit_Str_G_Max : LREAL;

//2025.01.04.131102 | 增加色组印长 -4字节
	rLength_Printing : REAL;		//色组印长 -4字节
(*2025.3.5.153256移植新的套色算法-增加150个字节786-636*)
	stStArc_Mol_Param	:StArc_Mol_Param;
//2025.03.14.181709 | 带长计算的滤波次数	---2字节
	iBandLengthFilterCnt			: INT;

	iCoefOfCoupling_V 	 :INT;
(*2025.3.21.195756||新增*)
	byFollowColorId				: BYTE;
	xWaitFilmLenth_Follow1U		: BOOL;
	wButtonFun_Lamp					:WORD ;(*HMI界面按钮及指示灯			*)
	wSwitchFun						:WORD ;(*界面开关*)

	//Filter原本的wRsv在这里改一下改为从站精采样数据低通滤波频率
	uilowpasscutoff_hz				:UINT;
//2025.11.7.142851先把数据统一了，dwSlaveBtn_HMI分两个word,一个暂时baoliu
//	dwSlaveBtn_HMI					:DWORD;(*界面按钮						*)
(* 2021.12.23.153801/hdp *)
	rLong_Step_Roller_Pressure					: REAL;(* 压力步进值-长步|MM *)
	rShort_Step_Roller_Pressure					: REAL;(* 压力步进值-短步|MM *)

	rSV_UnitTemCtl					:REAL ;(*加热设定温度					*)

(*原用户基础工艺开关控制位直接用BIT吧，不用dwCtlBits_UnitBaseCraft了--
通讯改为共用体吧*)
(*bit0-bit31--2025.8.13.100117*)
	xSwitch_ScraperAuto					: BIT;(*刮刀手自动-bit0*)
	xSwitch_ScraperOn					: BIT;(*刮刀开关bit1*)
	xInterver_ScraperRun				: BIT;(*刮刀开关bit2*)
	xRsv_BIT3							: BIT;(*BIT3预留*)
	xSwitch_InkRollerAuto				: BIT;(*递墨辊手自动bit4*)
	xSwitch_InkRollerCW					: BIT;(*递墨辊正转bit5*)
	xSwitch_InkRollerCCW				: BIT;(*递墨辊反转bit6*)
	xInterver_InkRollerRun				: BIT;(*递墨辊运行bit7*)
	xSwitch_HotWindOn					: BIT;(*热风开关bit8*)
	xInterver_HotWindRun				: BIT;(*热风1运行bit9*)
	xRsv_BIT10							: BIT;(*BIT10预留*)
	xRsv_BIT11							: BIT;(*BIT11预留*)
	xSwitch_HotWindOn_II				: BIT;(*热风开关bit12*)
	xInterver_HotWindRun_II				: BIT;(*热风1运行bit13*)
	xRsv_BIT14							: BIT;(*BIT14预留*)
	xRsv_BIT15							: BIT;(*BIT15预留*)
	xSwitch_HeatingMode_Water			: BIT;(*水加热开关bit16*)
	xSwitch_HeatingMode_Ele				: BIT;(*电加热开关bit17*)
	xSwitch_Heating_I					: BIT;(*加热I档bit18*)
	xSwitch_Heating_II					: BIT;(*加热II档bit19*)
	xSwitch_Heating_III					: BIT;(*加热III档bit20*)
	xRsv_BIT21							: BIT;(*BIT21预留*)
	xRsv_BIT22							: BIT;(*BIT22预留*)
	xErrReset_Scraper					: BIT;(*刮刀故障复位bit23*)
	xErrReset_InkRoller					: BIT;(*递墨故障复位bit24*)
	xErrReset_Hotwind					: BIT;(*热风故障复位bit25*)
	xErrReset_Hotwind_II				: BIT;(*热风2故障复位bit26*)
	xErrReset_ExhAir					: BIT;(*排风故障复位bit27*)
	xSwitch_ExhAir						: BIT;(*排风开关bit28*)
	xInterver_ExhAir					: BIT;(*排风运行bit29*)
	xRsv_BIT30							: BIT;(*BIT30预留*)
	xSwitch_Coolwind					: BIT;(*冷风开关*)
(*基础工艺开关-*)
	dwCtlBits_UnitBaseCraft					: DWORD;(* 用户基础工艺控制位/加热/递墨辊/刮刀/热风 *)
												(*
												/ .bit0 ~bit3  刮刀
												/	/.bit0 刮刀自动(TRUE)/手动(FALSE)
												/	/.bit1 刮刀开(TRUE)/关(FALSE)
												/	/.bit2 刮刀运行信号/控制变频器启动
												/	/.bit3
												/ .bit4 ~bit7  递墨辊
												/	/.bit4 递墨辊自动(TRUE)/手动(FALSE)
												/	/.bit5 递墨辊正转(TRUE)/关或反转(FALSE)
												/	/.bit6 递墨辊反转(TRUE)/关或正转(FALSE)
												/	/.bit7 递墨辊运行信号/控制变频器启动-与/.4/.5共同确定正转还是反转
												/ .bit8 ~bit11 热风I
												/	/.bit8 热风I开(TRUE)/关(FALSE)
												/	/.bit9 热风I运行信号/控制变频器启动
												/	/.bit10
												/	/.bit11
												/ .bit12~bit15 热风II
												/	/.bit12 热风II开(TRUE)/关(FALSE)
												/	/.bit13 热风II运行信号/控制变频器启动
												/	/.bit14
												/	/.bit15
												/ .bit16~bit23
												/	/ .bit16 加热方式（水）
												/	/ .bit17 加热方式（电）
												/	/ .bit18 I档
												/	/ .bit19 II档
												/	/ .bit20 III档
												/	/ .bit21
												/	/ .bit22
												/ .bit23~bit26
												/	/ .bit23 刮刀故障复位
												/	/ .bit24 递墨故障复位
												/	/ .bit25 热风I故障复位
												/	/ .bit26 热风II故障复位
												/   / .bit27 排风故障复位
												/ .bit28~bit31 /2022.3.23.152646/hdp/预分配好/为和界面作绑定
												/	/ .bit28 排风开(TRUE)/关(FALSE)
												/	/ .bit29 排风运行信号/控制变频器启动
												/	/ .bit30
												(*2022.4.20.091641 移动到此处*)
												/	/ .bit31: 2022.4.20.091632|冷风机开关使能位||
												*)
(* 递墨辊部分 *)
	rHz_UnitInkRoller_ManuallySet			: REAL;(* 递墨辊手动输入频率/0.00~100.00Hz/协议Mailbox直接传输 *)
	rCoeff_UnitInkRoller_Auto				: REAL;(* 递墨辊自动系数/Mailbox双向/主从可设置/ *)
(* 刮刀部分 *)
	rHz_UnitScraper_ManuallySet				: REAL;(* 刮刀手动输入频率/0.00~100.00Hz/协议Mailbox直接传输 *)
	rCoeff_UnitScraper_Auto					: REAL;(* 刮刀自动系数/Mailbox双向/主从可设置/ *)
(* 热风部分 *)
	rHz_UnitHotWind_ManuallySet				: REAL;(* 热风频率/Mailbox双向/主从可设置/ |修改了命名*)
(*2022.3.22.154047 增加*)
	rHz_UnitHotWind_2_ManuallySet			: REAL;(* 热风II频率 |修改了命名*)
(*2022.3.22.154031 增加的*)
(*E<<<<<<<<<<<<<<<<<<<<<<<<<<<<<<<<<<<<<<<<<<<<<<<<<<*)
	byHotBlower_AO							: BYTE;(*2025.6.14.100346*)
	wAirReturnWindDoorValue					: WORD;(* 回风口风门开度值|输入范围(0~100),默认值:0;|2018.11.27.140852|xie.gc重新修改定义| *)
	wAirExhaustWindDoorValue				: WORD;(* 排风口风门开度值|输入范围(0~100),默认值:0;|2018.11.27.140852|xie.gc重新修改定义| *)

	rGirth_Sam								: REAL;(*套色采样的周长*)
	uiNum_Sam								: UINT;(*套色采样的减速比分子*)
	uiDen_Sam								: UINT;(*套色采样的减速比分m母*)
	rHz_UnitExhaust_ManuallySet				: REAL;(* 排风频率/Mailbox双向/主从可设置/ *)

	(*光纤电眼控制相关变量*)
	bySignalSelect					:BYTE;(*光纤电眼信号选择		*)
	//xi.hy//新增
	rOffset_T1						:REAL;	//T1路光纤偏移
	rSource_Light_T1       			:REAL;  //T1路光纤光源
	rBias_T1			  			:REAL;  //T1路光纤电眼偏置
	rBrightness_Light_T1			:REAL;  //T1路光纤电眼亮度

	rOffset_T2						:REAL;  //T2路光纤偏移
	rSource_Light_T2				:REAL;  //T2路光纤光源
	rBias_T2						:REAL;  //T2路光纤电眼偏置
	rBrightness_Light_T2			:REAL;  //T2路光纤电眼亮度

	rK_ArcErr_Lp											: REAL;(*套色误差低通滤波处理的K值*)
	rFilmLengthFromPrevPressUnit							: REAL;(*从前一个合压色到当前色的料长@mm|1色是=0@还未实现呢2024.05.25.130043*)
	byAve_v_extra							: BYTE;(*界面误差显示平均值*)
	xWaitFilmLenth_FollowPreU:BOOL;(*等料长标志区分为等待前一色*)
	xWaitFilmLength					: BOOL;
	(*新增变量|wang.nt|2025.08.07.204018*)
	rStep_OfChangeGirth :REAL ;  (*涂布版轴修改步幅*)
	uiTimeMs_RollerPressUpKeep : UINT ;      (*压辊双气缸-离压保持时间*)
	//9905界面内容
	rAxisVelPrf_Coeff1 				: REAL;
	rAxisVelPrf_Coeff2 				: REAL;
	rAxisVelPrf_Coeff3 				: REAL;
	rMargin_Mag_Arc 				: REAL;
	rMargin_Phi_Arc 				: REAL;
	rKp_MolCal 						: REAL;
	rKi_MolCal 						: REAL;
	byCompensateValue_Hor 			: BYTE;
	byMaxAddValue_Total_Hor 		: BYTE;
	rWn_Arc 						: REAL;
	rBw_Arc 						: REAL;
	rDp_Arc 						: REAL;
	rK 								: REAL;
	rA2 							: REAL;
	rA1 							: REAL;
	rA0 							: REAL;
	rG_Periodic 					: REAL;
	rW_Periodic 					: REAL;
	byCnt_Comm2ARM					: BYTE;

	(*2025.8.9.141718|部分位变量处理*)
	xBtnLinkage_HMI			: BIT;(*界面联动按钮*)
	xFlag_InkRollerRisen	: BIT;(*递墨辊升起标志*)
	(*新增变量-开始|wang.nt2025.08.13.165332*)
	xInValidVirtualCnt:BOOL;(*虚拟马盘非法值*)
	byBrakeResistanceAlarm:byte;
	(*新增变量-结束|wang.nt2025.08.13.165332*)
	(*新增工艺参数|2025.08.15.151930*)
	byFreq_ExhaustAir  : BYTE ;
	byAirInletWindDoorValue : BYTE ;
	(*新增等料长相关参数|2025.08.20.214206*)
	lrPreReg_ConstVal						: LREAL;(*预套准色组间固定料长部分|单位:mm*)
	//xSkipHeaderSts							: BOOL;(*让料头状态@每次接料都会计算@根据是否打开让料头标志是否输出xSkipHeader*)
	//xSkipHeader								: BOOL;(*让料头*)
	(*预套准相关变量|wang.nt|2025.08.21.162244*)
	uiTurnOverFilmLenth						: UINT;(*翻料架料膜长度@mm*)
	iPhase_Locating						: INT;(*固定相位|2024.9.25.174406|Wang.nt*)
	iPhase_RegisterOk						: INT;(*套准相位|版套印准确的相位<通用相位和相位保存/恢复都可以复用该变量>|*)
	iPhase_FinalUsed						: INT;(*通用相位-最终用相位|*)
	iPhase_InstallPlate						: INT;(*装版相位|*)
	byPhaseState:BYTE;(*/.0 数值有效无效位|./1 数据需要保存标志位|/.4更新成功了|/.5 更新失败了*)(*马克线位置处理-世标*)
	xPreRegisterValid_Manu					: BOOL;(*手动预套有效*)
	iStationId								: INT;(*对应的站号|每次开机和更新系统配置都会重新更新的*)
	xServoOn								: BOOL;(*伺服使能|调用过GT_AxisOn就会被置位,GT_AxisOff会被清除*)
	lrPT_Pos								: LREAL;(*轴PT位置|*)
	diPT_Time								: DINT;(*轴PT时间值|*)
	iPT_Type								: INT;(*轴PT段选择|PT_SEGMENT_NORMAL;PT_SEGMENT_EVEN*)
	xPT_DataValid							: BOOL;(*轴PT数据有效|*)
	wEnableMode_Motor						: WORD;
	byFakeThreshold_V				:BYTE;(*纵向飞点阀值@丝			*)
	byFakeThreshold_H				:BYTE;(*横向飞点阀值@丝			*)
	byOvensAirOutWindDoorValue	: BYTE;
	xSwitch_TempFromEnc_PT1000							: BIT;
	xSwitch_MotorTemp_PT1000_NTC						: BIT;
//2025.12.30.222558新增变量，数据大小变化
(*2022.4.22.114421 排风风门变量添加|10bytes*)
	xUnitExhaustDamperCtl_Auto				: BOOL;(*排风风门控制自动*)
	rUnitExhaustDamperPos_ManuallySet		: REAL;(*排风风门位置手动设置值*)
	rUnitExhaustDamperPos_Cur				: REAL;(*排风风门写入当前位置值*)
	//新增超旭026.02.05.164858
	wButtonAndSwitch_ChaoXu	: WORD;	//.0 匀墨
										//.1 网辊锁轴
										//.2 充气
										//.3 墨盘电磁阀升
										//.4 照明
										//.5 确认修改版周
										//.6
										//.7
										//.8
										//.9
										//.10
										//.11 合压
										//.12 离压
										//.13
										//.14

END_STRUCT
END_TYPE

{IMPLEMENTATION}
